(* IEC 61131-3 sources: daoli-st-library/DL_Motion (part 23) *)

(* ---- FB_DL_GantrySyncAxis.st ---- *)
(*==============================================================================
 * 组件名称 (Component)  : FB_DL_GantrySyncAxis
 * 所属子库 (Sublibrary) : DL_Motion
 * 当前版本 (Version)    : 1.0.0
 * 组件分类 (Category)   : 功能块（FUNCTION_BLOCK）· 多轴同步耦合族 · 龙门双驱偏斜保护
 * 兼容性   (Platform)   : CODESYS 3.5 / TwinCAT 3 / 汇川 InoProShop / Schneider
 *                         Machine Expert；仅依赖 Standard.library
 *                         （TON / R_TRIG / LIMIT / MIN / MAX / ABS），零厂商方言
 * 接口依赖 (Depends)    : I_DL_MotionAxis / E_DL_AxisState（既有契约，Round 05，零修改）
 * 功能描述 (Function)   : 双驱龙门同步与偏斜保护。主动侧（主轴）与从动侧（从轴）
 *                         1:1 速度耦合，实时监视两侧实际位置偏差；两级阈值（预警
 *                         / 故障）分别触发降速纠偏与双轴停止；可选比例纠偏（偏差
 *                         为正即主动侧在前 → 从动侧加速追赶）；任一轴故障同拍双轴
 *                         停止（不对称风险优先，不做「健康侧继续」策略）。
 * 设计要点 (Key notes)  :
 *   ① 两级监视是本块骨架：预警阈只告警与纠偏，故障阈才双停；预警阈必须小于
 *      故障阈，组态写反时自动对调并提示（沿用库内对调自修复先例）。
 *   ② 偏差确认走延时（抗单拍毛刺）；延时参数变化时显式断输入一拍，使已计时
 *      归零（防「改时间常数后计时不清零」的幽灵故障）。
 *   ③ 纠偏为比例律 + 修正量限幅，不用积分（避免在轴外层再套积分器造成饱和）；
 *      长时间饱和判为机械卡滞或增益不足，升为故障级锁存。
 *   ④ 偏差回差 80% 才退出纠偏态，防止阈值边缘反复抖动。
 * 开源溯源 (Origin)     : 原创实现，clean-room。语义来源为公开技术文章「双编码器
 *                         龙门组态」（两级位置差监视、偏差锁存门限）、公开厂商
 *                         帮助的软龙门章节（两级监视：一级可复位、二级不可复位）、
 *                         公开论文「宽跨距龙门吊防偏斜控制器」（偏差 → 速度修正
 *                         量、增益限幅）与公开的数控龙门位置公差参考值（来源编号
 *                         RAW_NOTES S-3）。
 *                         「借鉴对象的许可说明」：上述对象均为公开发布但受版权
 *                         保护的帮助文档 / 技术文章 / 公开论文，属「可免费查阅、
 *                         仅借鉴语义与参数域」类别；本实现未复制任何源码或组态
 *                         文件，状态机、引脚命名、故障码与对调自修复策略均为本
 *                         库自有设计。
 * 验收向量 (Acceptance) :
 *   V1 正常耦合：使能后进入 eRun，偏差在预警阈内 → bInSync 为 TRUE；
 *   V2 注入 1 mm 偏差：进入 eCorrecting，修正量不超上限，偏差收敛后回 eRun；
 *   V3 偏差 3 mm（超故障阈 2 mm）持续 60 ms：确认后双轴同时停止 + 锁存 0273；
 *   V4 单轴故障：同拍双轴停止 + 锁存 0274（不等待偏差阈值）；
 *   V5 阈值写反（预警 5 / 故障 1）：自动对调 + 信息级 0151，仍能正常监视；
 *   V6 纠偏饱和持续 3 s：锁存 0271；
 *   V7 偏差未回到预警阈内给 bReset：拒绝复位 + 信息级 0150；
 *   V8 位置含非有限值：锁存 0272 并立即双停；
 *   V9 运行中途插入跟踪脉冲 bTrack：清偏差计时、退回 eIdle（公约 0.1）。
 * 已知限制 (Limits)     :
 *   ① 本块为逻辑层同步监视与纠偏编排，不构成 ISO 13849 / IEC 62061 认证安全
 *      功能；机械偏斜的最终保护由硬件限位与安全回路承担。
 *   ② 两侧轴若注入同一实例，块内无法识别，轴自身仲裁；调用方须保证主动侧与
 *      从动侧为不同实例。
 *   ③ 偏差延时确认粒度等于任务扫描周期，极短延时（小于两个扫描周期）实际等效
 *      单拍确认，毛刺风险由调用方通过 tDevDelay 规避。
 * 规格偏离 (Deviation)  :
 *   ① 依公约 0.1 增补 bTrack 输入引脚（首扫 / 跟踪范式强制项）。
 *   ② 进入 eStopping 后沿用本块既有的停止单发标志，避免每拍重复下发停止指令；
 *      规格「同拍对两轴各发一次」在进入该态的同一拍内完成，语义不变。
 *   ③ 使能撤除时在清零输出的同时补发一次双轴停止（安全保守处置）。
 *   ④ 故障级码 0270（阈值非法）在使能期间逐拍复核，一旦组态被改坏立即锁存，
 *      不停留在仅启动时校验。
 * 红线自检 (Redline)    :
 *   R1 零全局符号区访问 ✓（无全局变量表访问、无外部变量声明）
 *   R2 零物理地址直写 ✓（无输入输出通道地址记号）
 *   R3 纯 IEC 61131-3 ✓（仅 TON / R_TRIG / LIMIT / MIN / MAX / ABS）
 *   R4 防除零 / 防越界 / 浮点容差 ✓（阈值对调与回差全用容差比较、无数组索引、
 *      时间参数变化断输入一拍）
 *   R5 声明行 100% 中英双语同行注释 ✓
 *   R6 ENUM + CASE 且 CASE 含 ELSE 兜底 ✓
 *   R7 定时器与边沿实例无条件周期刷新 ✓（本块无单拍脉冲输出）
 *   POU 终结符成对 ✓（FUNCTION_BLOCK ↔ END_FUNCTION_BLOCK，末行即终结符；
 *   TYPE ↔ END_TYPE 成对）
 * 故障码表 (Error codes):
 *   16#0004_0150【信息级】偏差未回预警阈内，复位被拒；
 *   16#0004_0151【信息级】预警 / 故障阈值对调自修复；
 *   16#0004_0152【信息级】纠偏速度上限非法回默认；
 *   16#0004_0270【故障级】偏差阈值非法（≤0 / 非有限值），锁存；
 *   16#0004_0271【故障级】纠偏长时间饱和（疑似机械卡滞），锁存；
 *   16#0004_0272【故障级】轴位置信号非有限值，锁存；
 *   16#0004_0273【故障级】偏差超故障阈触发双轴停止，锁存；
 *   16#0004_0274【故障级】单轴故障触发双轴停止（透传），锁存；
 *   16#0004_0297【故障级】非法状态兜底（本块专用，不与其他块共用）。
 *   信息级码只进 uErrorId；bFault 为派生式仅反映 eFault 态。
 * 修订历史 (Revision)   :
 *   2026-11-15  v1.0.0  首版入库（Round 08 · DL_Motion 同步耦合族）
 *============================================================================*)

(*-----------------------------------------------------------------------------
 * 调用示例 (Instance guide)：
 *   fbGantry.iMasterAxis := fbLeftAxis;           // 主动侧（驱动侧）实例
 *   fbGantry.iSlaveAxis  := fbRightAxis;          // 从动侧（跟随侧）实例
 *   fbGantry(bEnable := bGantryOn,
 *            fDevTolWarn := 0.5, fDevTolFault := 2.0,
 *            tDevDelay := T#50MS, bCorrectEnable := TRUE,
 *            fCorrGain := 2.0, fCorrSpeedMax := 20.0,
 *            fCoupleSpeed := 10.0, fAcc := 500.0);
 *   IF fbGantry.bStopBothCmd THEN bSafetyRelayDrop := TRUE; END_IF
 *   注：两侧轴的上使能、回原与限位保护仍由各自轴块与安全链负责，本块只做
 *       速度耦合与偏差监视。
 *----------------------------------------------------------------------------*)

(*-----------------------------------------------------------------------------
 * 常见误用与现场提示 (Field notes)：
 *   1 预警阈与故障阈不要设成同值：同值时监视失去两级意义，块内会按对调处理
 *      并提示，但工艺上应重新组态（预警阈建议取故障阈的 1/4 ~ 1/2）。
 *   2 纠偏增益过大会在阈值边缘产生速度抖动；从 1.0 ~ 3.0 起步，观察
 *      fCorrSpeedCmd 是否长期贴上限（贴上限即增益不足或机械卡滞）。
 *   3 单轴报跟随误差时本块同拍双停，另一轴不会「继续跑」——这是刻意的保守
 *      策略，复位后必须人工确认横梁已回正再重新使能。
 *   4 bFault 一旦置位只能靠 bReset 上升沿解除，且要求偏差已回到预警阈内；
 *      机械偏斜未消除时复位会被拒（信息级 0150），必须先手动点动纠偏。
 *   5 本块不产生位置指令，只产生速度指令；位置同步精度取决于两侧驱动自身
 *      的位置环，本块不替代驱动的位置控制。
 *   6 阈值组态被改坏（≤0 / 非有限值 / 超域）时本块直接锁存 0270，且「组态未改好
 *      之前复位会立刻再次锁存」是刻意行为：不允许带着非法偏差阈值运行龙门。
 *----------------------------------------------------------------------------*)

(*-----------------------------------------------------------------------------
 * 枚举: E_DL_GantryState（归属 DL_Motion，与本功能块同文件发布）
 * 含义: 龙门双驱同步状态机，编号间隔 10 预留扩展位。
 *----------------------------------------------------------------------------*)
{attribute 'strict'}
{attribute 'qualified_only'}
TYPE E_DL_GantryState :
(
    eIdle       := 0,    // 空闲：未耦合，输出全清 / Idle: not coupled, outputs cleared
    eCoupling   := 10,   // 耦合建立：双轴以慢速趋同 / Coupling: both axes converge at low speed
    eRun        := 20,   // 运行：1:1 速度跟随 + 偏差监视 / Run: 1:1 velocity follow with deviation monitoring
    eCorrecting := 30,   // 纠偏中：偏差超预警阈且纠偏使能 / Correcting: deviation over warn band with correction enabled
    eStopping   := 40,   // 双轴停止中：偏差超故障阈或任一轴故障 / Stopping: deviation over fault band or axis fault
    eFault      := 99    // 故障锁存：仅 bReset 上升沿且偏差回位可退出 / Fault: latched, bReset only after deviation recovered
) UINT;
END_TYPE

FUNCTION_BLOCK FB_DL_GantrySyncAxis
VAR_INPUT
    bEnable         : BOOL := FALSE;        // 总使能（Enable），FALSE=停止并清指令，电平语义
    bReset          : BOOL := FALSE;        // 复位故障（Reset），上升沿受理，须偏差已回预警阈内才真正复位
    bTrack          : BOOL := FALSE;        // 偏差计时重同步（Tracking pulse），上升沿即清计时与锁存并退回 eIdle
    fDevTolWarn     : REAL := 0.5;          // 偏差预警阈（Deviation warn tolerance）[mm]，域 0.001..50，须小于故障阈
    fDevTolFault    : REAL := 2.0;          // 偏差故障阈（Deviation fault tolerance）[mm]，域 0.01..100
    tDevDelay       : TIME := T#50MS;       // 偏差确认延时（Deviation confirm delay）[ms]，超阈须持续此时间才动作
    bCorrectEnable  : BOOL := TRUE;         // 纠偏使能（Correction enable），FALSE=只监视不纠偏
    fCorrGain       : REAL := 2.0;          // 纠偏比例增益（Correction gain）[1/s]，域 0..50，0=纠偏关闭
    fCorrSpeedMax   : REAL := 20.0;         // 纠偏速度修正上限（Correction speed limit）[mm/s]，域 0.1..500
    fCoupleSpeed    : REAL := 10.0;         // 耦合建立慢速（Coupling speed）[mm/s]，域 0.1..1000，双轴以此速度趋同
    fAcc            : REAL := 500.0;        // 加/减速度（Acceleration）[mm/s²]，域 0.1..100000，非有限值回默认
END_VAR
VAR_OUTPUT
    bInSync         : BOOL := FALSE;        // 同步中（In sync），eRun / eCorrecting 且偏差未超预警阈为 TRUE
    fDeviation      : REAL := 0.0;          // 实时偏差（Deviation）[mm]，= 主动侧位置 − 从动侧位置，带符号
    bDevWarn        : BOOL := FALSE;        // 偏差预警（Deviation warning），延时确认后置位，回差内自动清，瞬态型
    bFault          : BOOL := FALSE;        // 故障锁存（Fault），派生式仅故障级码参与，信息级码不置位
    uErrorId        : UDINT := 0;           // 故障码（Error code），段位 16#0004_xxxx，0=无故障
    bStopBothCmd    : BOOL := FALSE;        // 双轴停止请求（Stop both request），供上层安全链与 HMI 监视
    fCorrSpeedCmd   : REAL := 0.0;          // 纠偏速度修正量（Correction speed）[mm/s]，带符号，叠加到从动侧指令
END_VAR
VAR_IN_OUT
    iMasterAxis     : I_DL_MotionAxis;      // 主动侧轴接口引用（Drive side axis），由调用方注入
    iSlaveAxis      : I_DL_MotionAxis;      // 从动侧轴接口引用（Following side axis），由调用方注入
END_VAR
VAR
    eState          : E_DL_GantryState := E_DL_GantryState.eIdle; // 内部状态机步序（Internal state）
    bInit           : BOOL := FALSE;        // 首扫完成标志（First-scan done flag），初值 FALSE，随 bTrack 复位
    bFaultLatch     : BOOL := FALSE;        // 故障锁存标志（Fault latch），仅 bReset 沿或新啮合沿解除
    bRefOk          : BOOL := FALSE;        // 双引用有效标志（Both references valid），逐拍重算
    bStopIssued     : BOOL := FALSE;        // 双轴停止已下发标志（Stop issued flag），单发化防重复发令
    bWarnLatched    : BOOL := FALSE;        // 预警锁存标志（Warning latched），带回差自动清除
    bMonActive      : BOOL := FALSE;        // 偏差监视使能（Monitoring active），运行三态为 TRUE
    bParamBad       : BOOL := FALSE;        // 阈值参数非法标志（Tolerance parameter invalid），逐拍重算
    bDelayChanged   : BOOL := FALSE;        // 延时参数变更标志（Delay changed flag），断输入一拍用
    fWarnEff        : REAL := 0.5;          // 生效预警阈（Effective warn tolerance）[mm]，对调后值
    fFaultEff       : REAL := 2.0;          // 生效故障阈（Effective fault tolerance）[mm]，对调后值
    fCorrMaxEff     : REAL := 20.0;         // 生效纠偏上限（Effective correction limit）[mm/s]，非法回默认
    fAccEff         : REAL := 500.0;        // 生效加减速度（Effective acceleration）[mm/s²]，非法回默认
    fCoupleEff      : REAL := 10.0;         // 生效耦合慢速（Effective coupling speed）[mm/s]，非法回默认
    fDevAbs         : REAL := 0.0;          // 偏差绝对值（Absolute deviation）[mm]，阈值比较用
    fCorrAbs        : REAL := 0.0;          // 纠偏量绝对值（Absolute correction）[mm/s]，饱和判定用
    fCorrCmd        : REAL := 0.0;          // 纠偏修正量（Correction command）[mm/s]，带符号
    fMasterPos      : REAL := 0.0;          // 主动侧位置（Drive side position）[mm]
    fSlavePos       : REAL := 0.0;          // 从动侧位置（Following side position）[mm]
    fMasterVel      : REAL := 0.0;          // 主动侧速度（Drive side velocity）[mm/s]，带符号
    fSlaveVel       : REAL := 0.0;          // 从动侧速度（Following side velocity）[mm/s]，带符号
    fCmdVel         : REAL := 0.0;          // 下发给从动侧的速度指令（Commanded velocity）[mm/s]，带符号
    tDelayEff       : TIME := T#50MS;       // 生效确认延时（Effective confirm delay）[ms]，负值归零
    tDelayPrev      : TIME := T#0MS;        // 上拍确认延时（Previous confirm delay）[ms]，变更检测基准
    nStopCode       : UDINT := 0;           // 停止原因码（Stop reason code），进 eFault 时落地
    fbTrigReset     : R_TRIG;               // 复位指令上升沿（Reset command rising edge）
    fbTonDevWarn    : TON;                  // 偏差预警延时确认（Warn confirm delay timer）
    fbTonDevFault   : TON;                  // 偏差故障延时确认（Fault confirm delay timer）
    fbTonCorrSat    : TON;                  // 纠偏饱和累计计时（Correction saturation timer）
END_VAR
VAR CONSTANT
    DL_GANTRY_INF_MAX   : REAL := 1.0E30;   // 有限值判定幅值上限（Finite magnitude bound）[无量纲，按比较量量纲同值使用]
    DL_GANTRY_EPS       : REAL := 1.0E-6;   // 浮点判零容差（Float zero tolerance）[无量纲，按比较量量纲同值使用]
    DL_GANTRY_TOL_MIN   : REAL := 1.0E-3;   // 阈值下限（Tolerance floor）[mm]，低于此值判非法
    DL_GANTRY_TOL_MAX   : REAL := 100.0;    // 阈值上限（Tolerance ceiling）[mm]，高于此值判非法
    DL_GANTRY_CORR_DEF  : REAL := 20.0;     // 纠偏上限默认值（Default correction limit）[mm/s]
    DL_GANTRY_CORR_MAX  : REAL := 500.0;    // 纠偏上限允许最大值（Correction limit ceiling）[mm/s]
    DL_GANTRY_ACC_DEF   : REAL := 500.0;    // 加速度默认回退值（Default acceleration）[mm/s²]
    DL_GANTRY_CPL_DEF   : REAL := 10.0;     // 耦合慢速默认回退值（Default coupling speed）[mm/s]
    DL_GANTRY_HYST      : REAL := 0.8;      // 回差系数（Hysteresis factor）[-]，低于预警阈 80% 才清预警
    DL_GANTRY_SAT_RATIO : REAL := 0.98;     // 饱和判定比例（Saturation ratio）[-]，达上限 98% 视为饱和
    DL_GANTRY_SAT_TIME  : TIME := T#3S;     // 饱和持续上限（Saturation time limit）[ms]，超过判卡滞
    DL_GANTRY_SPEED_BAND: REAL := 1.0E-5;   // 速度趋同判定带（Speed convergence band）[mm/s]，= 判零容差 × 10
    DL_GANTRY_ZERO_TIME : TIME := T#0S;     // 零延时字面量（Zero delay literal）[ms]，用于延时下限比较
END_VAR

// 段 1｜边沿实例无条件周期刷新（红线 R7：严禁置于 IF / CASE 分支内）
fbTrigReset(CLK := bReset);

// 段 2｜出口默认赋值（公约 0.9：早退路径输出必须确定）
bInSync       := FALSE;
bDevWarn      := FALSE;
bFault        := (eState = E_DL_GantryState.eFault);
fCorrSpeedCmd := 0.0;
fDeviation    := 0.0;

// 段 3｜双引用有效性判定 + 反馈量采集（无效时全部回零，定时器照样刷新）
bRefOk := (iMasterAxis <> 0) AND (iSlaveAxis <> 0);
IF bRefOk THEN
    fMasterPos := iMasterAxis.fPosition;
    fSlavePos  := iSlaveAxis.fPosition;
    fMasterVel := iMasterAxis.fVelocity;
    fSlaveVel  := iSlaveAxis.fVelocity;
ELSE
    fMasterPos := 0.0;
    fSlavePos  := 0.0;
    fMasterVel := 0.0;
    fSlaveVel  := 0.0;
END_IF
fDeviation := fMasterPos - fSlavePos;
fDevAbs    := ABS(fDeviation);

// 段 4｜阈值参数防御：非有限值 / 超域判非法，预警阈不小于故障阈时自动对调
fWarnEff  := fDevTolWarn;
fFaultEff := fDevTolFault;
bParamBad := FALSE;
IF (fWarnEff <> fWarnEff) OR (ABS(fWarnEff) > DL_GANTRY_INF_MAX)
   OR (fWarnEff < DL_GANTRY_TOL_MIN) OR (fWarnEff > DL_GANTRY_TOL_MAX) THEN
    bParamBad := TRUE;
END_IF
IF (fFaultEff <> fFaultEff) OR (ABS(fFaultEff) > DL_GANTRY_INF_MAX)
   OR (fFaultEff < DL_GANTRY_TOL_MIN) OR (fFaultEff > DL_GANTRY_TOL_MAX) THEN
    bParamBad := TRUE;
END_IF
IF (NOT bParamBad) AND (fWarnEff > (fFaultEff - DL_GANTRY_EPS)) THEN
    fWarnEff  := fDevTolFault;                           // 自动对调：写反时按对调后值监视，不静默
    fFaultEff := fDevTolWarn;
    uErrorId  := 16#0004_0151;                           // 【信息级】预警 / 故障阈值对调自修复
END_IF

IF (fCorrSpeedMax <> fCorrSpeedMax) OR (ABS(fCorrSpeedMax) > DL_GANTRY_INF_MAX)
   OR (fCorrSpeedMax < DL_GANTRY_TOL_MIN) THEN
    fCorrMaxEff := DL_GANTRY_CORR_DEF;                   // 纠偏上限非法 → 默认 20 mm/s
    uErrorId    := 16#0004_0152;                         // 【信息级】纠偏速度上限非法回默认
ELSE
    fCorrMaxEff := MIN(fCorrSpeedMax, DL_GANTRY_CORR_MAX);
END_IF

IF (fAcc <> fAcc) OR (ABS(fAcc) > DL_GANTRY_INF_MAX) OR (fAcc < DL_GANTRY_TOL_MIN) THEN
    fAccEff := DL_GANTRY_ACC_DEF;
ELSE
    fAccEff := fAcc;
END_IF

IF (fCoupleSpeed <> fCoupleSpeed) OR (ABS(fCoupleSpeed) > DL_GANTRY_INF_MAX) OR (fCoupleSpeed < DL_GANTRY_TOL_MIN) THEN
    fCoupleEff := DL_GANTRY_CPL_DEF;
ELSE
    fCoupleEff := fCoupleSpeed;
END_IF

// 段 5｜确认延时防御与变更检测（公约 0.6：语义参数变化必须断输入一拍）
IF tDevDelay < DL_GANTRY_ZERO_TIME THEN
    tDelayEff := DL_GANTRY_ZERO_TIME;                    // 负延时归零，按单拍确认（毛刺风险由调用方规避）
ELSE
    tDelayEff := tDevDelay;
END_IF
bDelayChanged := (tDelayEff <> tDelayPrev);              // 延时变更：本拍强制断输入，使已计时归零
tDelayPrev    := tDelayEff;

// 段 6｜偏差监视使能（运行三态参与监视）
bMonActive := (eState = E_DL_GantryState.eCoupling) OR (eState = E_DL_GantryState.eRun)
              OR (eState = E_DL_GantryState.eCorrecting);

// 段 7｜定时器无条件周期刷新（红线 R7：严禁置于 IF / CASE 分支内）
fbTonDevWarn(IN := bRefOk AND bMonActive AND (fDevAbs >= fWarnEff) AND (NOT bDelayChanged),
             PT := tDelayEff);
fbTonDevFault(IN := bRefOk AND bMonActive AND (fDevAbs >= fFaultEff) AND (NOT bDelayChanged),
              PT := tDelayEff);
fbTonCorrSat(IN := (eState = E_DL_GantryState.eCorrecting) AND (fCorrAbs >= fCorrMaxEff * DL_GANTRY_SAT_RATIO),
             PT := DL_GANTRY_SAT_TIME);

// 段 8｜引用无效直接退出（定时器已在上方无条件刷新，本拍不产生任何轴动作）
IF NOT bRefOk THEN
    RETURN;
END_IF

// 段 9｜预警锁存与回差清除（瞬态型，每拍重算）
IF fDevAbs >= fWarnEff THEN
    bWarnLatched := fbTonDevWarn.Q;                      // 超阈值区间：以延时确认结果为准
ELSIF fDevAbs <= (fWarnEff * DL_GANTRY_HYST) THEN
    bWarnLatched := FALSE;                               // 回差内自动清除
END_IF

// 段 10｜首扫与跟踪范式（公约 0.1：bTrack OR (NOT bInit) 为唯一判据，禁止反序）
IF bTrack OR (NOT bInit) THEN
    bWarnLatched := FALSE;
    bStopIssued  := FALSE;
    bStopBothCmd := FALSE;
    fCorrCmd     := 0.0;
    fCorrAbs     := 0.0;
    nStopCode    := 0;
    eState       := E_DL_GantryState.eIdle;
    bInit        := TRUE;                                // 首扫完成后置位（判据恒为 bTrack OR NOT bInit）
END_IF

// 段 11｜总使能撤除：清指令 + 补发一次双轴停止（安全保守处置）
IF NOT bEnable THEN
    IF (NOT bStopIssued) AND ((eState = E_DL_GantryState.eCoupling) OR (eState = E_DL_GantryState.eRun)
       OR (eState = E_DL_GantryState.eCorrecting)) THEN
        iMasterAxis.Stop();                              // 主动侧停止（本拍唯一一次主动侧调用）
        iSlaveAxis.Stop();                               // 从动侧停止（本拍唯一一次从动侧调用）
        bStopIssued := TRUE;
    END_IF
    eState    := E_DL_GantryState.eIdle;
    fCorrCmd  := 0.0;
    fCorrAbs  := 0.0;
END_IF

// 段 12｜事件码管理（公约 0.7 / R15）：锁存码仅在解除路径清，瞬时码逐拍重算
IF NOT bFaultLatch THEN
    uErrorId := 0;
END_IF

// 段 13｜位置 / 力矩类信号非有限值拦截（判定不可信，立即转双停）
IF (fMasterPos <> fMasterPos) OR (fSlavePos <> fSlavePos)
   OR (ABS(fMasterPos) > DL_GANTRY_INF_MAX) OR (ABS(fSlavePos) > DL_GANTRY_INF_MAX) THEN
    IF (eState <> E_DL_GantryState.eIdle) AND (eState <> E_DL_GantryState.eFault) THEN
        nStopCode := 16#0004_0272;                       // 【故障级】轴位置信号非有限值
        eState    := E_DL_GantryState.eStopping;
    END_IF
END_IF

// 段 14｜阈值非法拦截（使能期间逐拍复核组态）
IF bParamBad THEN
    IF eState <> E_DL_GantryState.eFault THEN
        bFaultLatch := TRUE;
        uErrorId    := 16#0004_0270;                     // 【故障级】偏差阈值非法
        eState      := E_DL_GantryState.eFault;
    END_IF
END_IF

// 段 15｜主状态机（ENUM + CASE + ELSE 兜底）
CASE eState OF

    E_DL_GantryState.eIdle:                              // 空闲：等待使能
        bInSync  := FALSE;
        bStopIssued := FALSE;
        bStopBothCmd := FALSE;
        fCorrCmd := 0.0;
        IF bEnable AND (NOT bParamBad) THEN
            bFaultLatch := FALSE;                        // 使能上升：锁存码解除路径（R15）
            fCorrCmd    := 0.0;
            eState      := E_DL_GantryState.eCoupling;
        END_IF

    E_DL_GantryState.eCoupling:                          // 耦合建立：双轴以慢速趋同
        bStopBothCmd := FALSE;
        IF iMasterAxis.bError OR iSlaveAxis.bError THEN
            nStopCode := 16#0004_0274;                   // 【故障级】单轴故障（不对称风险优先）
            eState    := E_DL_GantryState.eStopping;
        ELSIF fbTonDevFault.Q THEN
            nStopCode := 16#0004_0273;                   // 【故障级】偏差超故障阈
            eState    := E_DL_GantryState.eStopping;
        ELSE
            // 跟随主动侧速度，但幅值不超过耦合慢速
            fCmdVel := LIMIT(-fCoupleEff, fMasterVel, fCoupleEff);
            IF NOT iSlaveAxis.MoveVelocity(fVel := fCmdVel, fAcc := fAccEff) THEN
                bFaultLatch := TRUE;
                uErrorId    := 16#0004_0274;             // 【故障级】从动侧速度指令被拒（按单轴故障处置）
                eState      := E_DL_GantryState.eFault;
            ELSIF (ABS(fMasterVel - fSlaveVel) <= DL_GANTRY_SPEED_BAND) AND (fDevAbs <= fWarnEff) THEN
                eState := E_DL_GantryState.eRun;         // 速度趋同且偏差在预警阈内 → 运行
            END_IF
        END_IF

    E_DL_GantryState.eRun:                               // 运行：1:1 跟随，纠偏量为零
        IF iMasterAxis.bError OR iSlaveAxis.bError THEN
            nStopCode := 16#0004_0274;
            eState    := E_DL_GantryState.eStopping;
        ELSIF fbTonDevFault.Q THEN
            nStopCode := 16#0004_0273;
            eState    := E_DL_GantryState.eStopping;
        ELSE
            fCorrCmd := 0.0;                             // 运行态不纠偏
            IF bCorrectEnable AND (ABS(fCorrGain) > DL_GANTRY_EPS) AND bWarnLatched THEN
                eState := E_DL_GantryState.eCorrecting;  // 偏差确认超预警阈且纠偏使能 → 纠偏
            END_IF
            fCmdVel := fMasterVel;
            IF NOT iSlaveAxis.MoveVelocity(fVel := fCmdVel, fAcc := fAccEff) THEN
                bFaultLatch := TRUE;
                uErrorId    := 16#0004_0274;             // 【故障级】从动侧速度指令被拒
                eState      := E_DL_GantryState.eFault;
            END_IF
        END_IF

    E_DL_GantryState.eCorrecting:                        // 纠偏中：比例律修正量限幅
        IF iMasterAxis.bError OR iSlaveAxis.bError THEN
            nStopCode := 16#0004_0274;
            eState    := E_DL_GantryState.eStopping;
        ELSIF fbTonDevFault.Q THEN
            nStopCode := 16#0004_0273;
            eState    := E_DL_GantryState.eStopping;
        ELSIF fbTonCorrSat.Q THEN
            bFaultLatch := TRUE;
            uErrorId    := 16#0004_0271;                 // 【故障级】纠偏长时间饱和（疑似卡滞 / 增益不足）
            eState      := E_DL_GantryState.eFault;
        ELSE
            // 偏差为正（主动侧在前）→ 从动侧加速追赶；为负则减速
            fCorrCmd := LIMIT(-fCorrMaxEff, fCorrGain * fDeviation, fCorrMaxEff);
            fCorrAbs := ABS(fCorrCmd);
            // 偏差回到预警阈 80% 以内（回差）→ 退出纠偏
            IF fDevAbs <= (fWarnEff * DL_GANTRY_HYST) THEN
                fCorrCmd := 0.0;
                fCorrAbs := 0.0;
                eState   := E_DL_GantryState.eRun;
            END_IF
            fCmdVel := fMasterVel + fCorrCmd;
            IF NOT iSlaveAxis.MoveVelocity(fVel := fCmdVel, fAcc := fAccEff) THEN
                bFaultLatch := TRUE;
                uErrorId    := 16#0004_0274;             // 【故障级】从动侧速度指令被拒
                eState      := E_DL_GantryState.eFault;
            END_IF
        END_IF

    E_DL_GantryState.eStopping:                          // 双轴停止：同拍各发一次，停稳后锁存
        bStopBothCmd := TRUE;
        fCorrCmd     := 0.0;
        fCorrAbs     := 0.0;
        IF NOT bStopIssued THEN
            iMasterAxis.Stop();                          // 主动侧停止（本拍唯一一次主动侧调用）
            iSlaveAxis.Stop();                           // 从动侧停止（本拍唯一一次从动侧调用）
            bStopIssued := TRUE;
        END_IF
        IF (ABS(fMasterVel) <= DL_GANTRY_EPS) AND (ABS(fSlaveVel) <= DL_GANTRY_EPS) THEN
            bFaultLatch := TRUE;
            IF nStopCode = 0 THEN
                uErrorId := 16#0004_0273;                // 【故障级】兜底：停止原因缺失时按偏差超限记账
            ELSE
                uErrorId := nStopCode;                   // 落地本次停止的真实原因码
            END_IF
            bStopIssued := FALSE;
            eState      := E_DL_GantryState.eFault;
        END_IF

    E_DL_GantryState.eFault:                             // 故障锁存：仅复位沿且偏差回位可退出
        bInSync      := FALSE;
        bStopBothCmd := TRUE;                            // 故障态保持停止请求，供安全链与 HMI 监视
        fCorrCmd     := 0.0;
        fCorrAbs     := 0.0;
        bStopIssued  := FALSE;
        IF fbTrigReset.Q THEN
            IF fDevAbs <= fWarnEff THEN
                bFaultLatch := FALSE;                    // 唯一解除路径：偏差已回预警阈内
                uErrorId    := 0;
                nStopCode   := 0;
                eState      := E_DL_GantryState.eIdle;
            ELSE
                uErrorId := 16#0004_0150;                // 【信息级】偏差未回预警阈内，复位被拒
            END_IF
        END_IF

    ELSE                                                 // 非法状态兜底（本块专用码）
        bFaultLatch  := TRUE;
        uErrorId     := 16#0004_0297;                    // 【故障级】非法状态兜底
        bInSync      := FALSE;
        bStopBothCmd := TRUE;
        fCorrCmd     := 0.0;
        fCorrAbs     := 0.0;
        eState       := E_DL_GantryState.eFault;

END_CASE

// 段 16｜出口映射（派生式，信息级码不参与 bFault）
bFault        := (eState = E_DL_GantryState.eFault);
bInSync       := ((eState = E_DL_GantryState.eRun) OR (eState = E_DL_GantryState.eCorrecting))
                 AND (NOT bWarnLatched);
bDevWarn      := bWarnLatched AND ((eState = E_DL_GantryState.eCoupling)
                 OR (eState = E_DL_GantryState.eRun) OR (eState = E_DL_GantryState.eCorrecting));
bStopBothCmd  := (eState = E_DL_GantryState.eStopping) OR (eState = E_DL_GantryState.eFault);
fDeviation    := fMasterPos - fSlavePos;
fCorrSpeedCmd := fCorrCmd;

END_FUNCTION_BLOCK

(* ---- FB_DL_LineInterp2Axis.st ---- *)
(*==============================================================================
 * 组件名称 (Component)  : FB_DL_LineInterp2Axis
 * 所属子库 (Sublibrary) : DL_Motion
 * 当前版本 (Version)    : 1.0.1
 * 组件分类 (Category)   : 功能块（FUNCTION_BLOCK）· 运动控制 · 两轴直线插补
 * 兼容性   (Platform)   : CODESYS 3.5 / TwinCAT 3 / 汇川 InoProShop / Schneider
 *                         Machine Expert；纯 IEC 61131-3（第 3 版）语法，
 *                         仅依赖 Standard.library（R_TRIG / SQRT / MIN / MAX / LIMIT）
 * 功能描述 (Function)   : 由起点、终点、合成速度与加速度生成两轴位置给定：单位向量分解、
 *                         单轴速度上限折算、梯形与三角速度曲线自适应、端点平滑减速、
 *                         暂停保持与故障保护。输出 X 与 Y 的位置给定、合成速度、完成度
 *                         与本次实际峰值速度。
 * 分层声明 (Layering)   : ① 本件只输出「位置给定」，不输出使能、回零与报警复位，也不直接
 *                         驱动物理轴——两轴的实际闭环由各自的单轴功能块承担，本件给出
 *                         给定值后由上层把给定接到单轴的相对或绝对运动接口；
 *                         ② 不读系统时钟、不读任务周期：插补时间增量由引脚注入，
 *                         保证结果可复现、跨平台一致；
 *                         ③ 不做圆弧与样条插补（属后续件），不做过象限与软限位判断
 *                         （软限位归运动层的软限位保护件）。
 * 周期纪律 (Cycle)      : 本件必须放在固定周期任务中调用，周期值通过标称周期引脚注入。
 *                         变周期任务（如带事件触发的任务）会直接造成速度与位置偏差，
 *                         因为时间增量按注入值推进、不按墙钟补偿。
 * 速度剖面 (Profile)    : 单侧加速度距离为合成速度平方除以两倍加速度；若两侧之和超过
 *                         路径总长则判为三角曲线，峰值速度降为「加速度乘路径长」的平方根，
 *                         加速距离取路径长的一半。临界相等（两侧之和恰等于路径长）按梯形
 *                         处理：此时峰值速度与期望合成速度相等，两种判法结果一致、不跳变。
 * 端点纪律 (Endpoint)   : 减速段出口强制把已走距离钳到路径总长，进度置 100，避免离散步长
 *                         越过终点导致给定超程；收尾速度保留峰值的若干比例，防止速度
 *                         指数衰减而出现「永远差最后一点」的爬行。
 * 开源溯源 (Origin)     : 来源标签 github-topics-motion。原创实现（参考 GitHub 运动控制与
 *                         结构化文本主题下开源运动库的共同形态：单位向量分解、合成速度
 *                         限幅、梯形与三角自适应三段结构；多份实现交叉印证其为社区共识
 *                         写法，非某一家独有）。速度剖面、临界判据、暂停策略、枚举、
 *                         状态机与全部码位 100% 本库独立设计，clean-room 实现，零代码行
 *                         复制。各上游仓库许可未逐条复核，按最严口径只借结构与参数域。
 * 依赖     (Depends)    : 无 DL_ 内部依赖；Standard.library: R_TRIG / SQRT / MIN / MAX / LIMIT
 * 故障码表 (Error codes):
 *   16#0004_0109【信息级】路径长度为零，当拍直接完成，给定等于起点
 *   16#0004_010A【信息级】标称周期越界已钳到 0.1 毫秒至 1 秒
 *   16#0004_010B【信息级】单轴速度上限参与折算，合成速度已被压低
 *   16#0004_010C【信息级】路径过短，速度曲线降为三角（无匀速段）
 *   16#0004_0204【故障级】速度、加速度、单轴限速或最大路径长参数非法（锁存）
 *   16#0004_0205【故障级】路径长度超过允许上限（锁存）
 *   16#0004_0206【故障级】输入含非有限值（NaN 或无穷），前置拦截（锁存）
 *   16#0004_0207【故障级】非法状态兜底（锁存，终端安全态）
 * 码位占用 (Slot)       : 信息级 0109 / 010A / 010B / 010C；故障级 0204 / 0205 / 0206 / 0207。
 *                         全部落在 R12 本件分配块内，无跨块借用、无段外哨兵值。
 * 拍序纪律 (Cycle order) :
 *   ① ePhase    ：段 7 状态机（唯一位移点），段 8 复位分支是唯一回退点
 *   ② fS 与 fV  ：只在加速、匀速、减速三段内推进；暂停段速度归零且不推进位移
 *   ③ _bDone    ：进入准备相与进入完成相两处写，互斥不覆盖
 *   ④ uErrorId  ：段 9 单一优先级链，全拍只写一次
 * 验收向量 (Acceptance) :
 *   V1 梯形：起点 0 0、终点 300 400 → 路径 500；速度 100、加速度 200、单轴限速 1000 →
 *      合成 100 未被压低、单侧加速距离 25，两侧 50 小于 500 判梯形，峰值 100；
 *      中点给定为 150 与 200、完成度 50、合成速度 100
 *   V2 单轴限速：与 V1 同参但 X 轴限速改为 50 → 折算 83.333，合成速度被压到 83.333，
 *      X 分量 83.333 乘 0.6 等于 50，恰好不超限
 *   V3 零长度：起终点相同 → 当拍完成、给定等于起点、进度 100、码 0109
 *   V4 临界：路径 50、单侧加速距离 25 → 和为 50 恰等于路径长，判梯形，峰值 100
 *   V5 三角：路径 40 → 两侧 50 大于 40 判三角，峰值 89.44、单侧加速距离 20
 *   V6 参数非法：加速度为 0 → 故障位置位、码 0204、忙碌为假
 * 偏离留档 (Deviation)  :
 *   ① 规格未规定暂停时的时间补偿策略，本件按「不做补偿」实现：恢复后从当前速度重新加速，
 *      但时间增量仍按标称周期推进，故暂停不会造成位置瞬跳。若需要恒速衔接，应在工艺层
 *      用缓停而非暂停。
 *   ② 规格的减速段出口只要求钳位，本件额外把进度强制置 100，避免浮点除法在末拍给出
 *      99.9999 而让画面闪烁。
 * 修订历史 (Revision)   :
 *   2026-11-15  v1.0.0  首版落盘（R12 · 泳道 C · 两轴直线插补件）
 *   2026-11-15  v1.0.1  终审修复两处：
 *                       ① 暂停恢复时速度阶跃——加速段出口只看「位移到加速距离」，恢复后
 *                       该条件当拍即成立，再加速被整段跳过，速度由零直接跳到峰值；
 *                       改为位移与速度双条件，并在恢复时按剩余距离分流到减速段。
 *                       ② 零长度路径的完成度与头注释矛盾（注释写 100、出口被覆写为 0），
 *                       完成相下补满值分支
 *============================================================================*)

(*------------------------------------------------------------------------------
 * 枚举: E_DL_LineInterpPhase（本块相位，归属本功能块并同文件发布）
 *       Phase enumeration owned by this block, one member per motion segment
 *-----------------------------------------------------------------------------*)
TYPE E_DL_LineInterpPhase :
(
    eIdle  := 0,   // 待机：等待启动沿，给定保持在起点 / Idle, waiting for the start edge
    ePrep  := 10,  // 准备：参数闸门、向量分解、速度剖面计算 / Preparation, the whole profile is computed here
    eAccel := 20,  // 加速：速度按加速度上升，位移按速度积分 / Acceleration segment
    eCruise:= 30,  // 匀速：速度保持峰值，位移按速度积分 / Constant speed segment
    eDecel := 40,  // 减速：速度按加速度下降，出口钳位到终点 / Deceleration segment
    eDone  := 50,  // 完成：完成标志保持，给定等于终点，等下一次启动 / Done, held until the next start
    eHeld  := 60,  // 暂停：速度归零、位移保持，恢复后重新加速 / Held, speed forced to zero
    eFault := 99   // 故障：参数或输入非法、路径超限、非法状态 / Fault, needs a reset to leave
);
END_TYPE

FUNCTION_BLOCK FB_DL_LineInterp2Axis
VAR_INPUT
    bEnable       : BOOL;                          // 使能，FALSE 时停止推进并回待机 [-] / Enable, stopping the move and returning to idle
    bReset        : BOOL;                          // 复位故障，上升沿有效 [-] / Rising edge clears the fault
    bStart        : BOOL;                          // 启动，上升沿有效（待机与完成态可受理）[-] / Rising edge starts the move in idle or done
    bHold         : BOOL;                          // 暂停，TRUE 时速度归零且位移保持 [-] / Pauses the interpolation while TRUE
    fStartX       : REAL;                          // 起点 X 坐标 [毫米] / Start X in millimetres
    fStartY       : REAL;                          // 起点 Y 坐标 [毫米] / Start Y in millimetres
    fEndX         : REAL;                          // 终点 X 坐标 [毫米] / End X in millimetres
    fEndY         : REAL;                          // 终点 Y 坐标 [毫米] / End Y in millimetres
    fPathSpeed    : REAL := 100.0;                 // 期望合成速度 [毫米每秒]，域大于 0 / Desired path speed, must exceed zero
    fAccel        : REAL := 500.0;                 // 加减速度 [毫米每二次方秒]，域大于 0 / Acceleration, must exceed zero
    fMaxSpeedX    : REAL := 1000.0;                // X 轴速度上限 [毫米每秒]，域大于 0 / X axis speed limit
    fMaxSpeedY    : REAL := 1000.0;                // Y 轴速度上限 [毫米每秒]，域大于 0 / Y axis speed limit
    fNominalCycle : REAL := 0.004;                 // 标称插补周期 [秒]，域 0.0001 到 1 / Nominal interpolation period
    fMaxPathLen   : REAL := 100000.0;              // 允许最大路径长度 [毫米]，域大于 0 / Maximum path length, must exceed zero
END_VAR
VAR_OUTPUT
    bBusy         : BOOL;                          // 插补进行中（含准备段）[-] / Interpolation running, preparation included
    bActive       : BOOL;                          // 位置给定有效（推进中或暂停中）[-] / Position command valid
    bDone         : BOOL;                          // 到达终点，保持到下一次启动 [-] / End reached, held until the next start
    fCmdX         : REAL;                          // X 位置给定 [毫米] / X position command
    fCmdY         : REAL;                          // Y 位置给定 [毫米] / Y position command
    fPathProgress : REAL;                          // 路径完成度 [百分之]，域 0 到 100 / Path progress in percent
    fPathVel      : REAL;                          // 当前合成速度 [毫米每秒] / Current path speed
    fPathLen      : REAL;                          // 本次路径总长 [毫米] / Total path length of this move
    fPeakVel      : REAL;                          // 本次实际峰值速度 [毫米每秒] / Effective peak speed of this move
    bError        : BOOL;                          // 故障级锁存，仅 0204 至 0207 置位 [-] / Latched fault, only fault level codes set it
    uErrorId      : UDINT;                         // 事件码，0 表示无事件 [代码] / Event code, zero means none
    eState        : E_DL_LineInterpPhase;          // 主状态机当前相位 [-] / Current phase of the main state machine
END_VAR
VAR
    fbTrigStart   : R_TRIG;                        // 启动沿检测，主周期无条件刷新 [-] / Start edge detector, refreshed unconditionally
    fbTrigReset   : R_TRIG;                        // 复位沿检测，主周期无条件刷新 [-] / Reset edge detector, refreshed unconditionally
    ePhase        : E_DL_LineInterpPhase := E_DL_LineInterpPhase.eIdle; // 内部相位，对外经 eState 输出 [-] / Internal phase exported as eState
    bInit         : BOOL := FALSE;                 // 首扫标志，初值 FALSE，判据取非 [-] / First-scan flag initialised FALSE
    bFaultLatch   : BOOL;                          // 故障锁存，仅复位分支清除 [-] / Fault latch, cleared by the reset path only
    uErrInt       : UDINT;                         // 故障级码寄存，锁存型 [代码] / Latched fault level code register
    uInfoCode     : UDINT;                         // 本拍信息级码，每拍重算 [代码] / Info level code recomputed every scan
    bDoneLatch    : BOOL;                          // 完成标志保持寄存器 [-] / Done hold register
    fDx           : REAL;                          // X 方向位移 [毫米] / X displacement
    fDy           : REAL;                          // Y 方向位移 [毫米] / Y displacement
    fLen          : REAL;                          // 路径长度 [毫米] / Path length
    fUx           : REAL;                          // X 单位向量分量 [无量纲] / X unit component
    fUy           : REAL;                          // Y 单位向量分量 [无量纲] / Y unit component
    fVEff         : REAL;                          // 生效合成速度 [毫米每秒] / Effective path speed
    fVLimit       : REAL;                          // 单轴限速折算后的合成速度上限 [毫米每秒] / Speed cap derived from axis limits
    fTmpX         : REAL;                          // X 轴限速折算中间量 [毫米每秒] / X cap temporary
    fTmpY         : REAL;                          // Y 轴限速折算中间量 [毫米每秒] / Y cap temporary
    fAccUse       : REAL;                          // 生效加速度 [毫米每二次方秒] / Effective acceleration
    fAccDist      : REAL;                          // 单侧加速距离 [毫米] / One-sided acceleration distance
    fPeak         : REAL;                          // 本次峰值速度 [毫米每秒] / Peak speed of this move
    fVDecelFloor  : REAL;                          // 收尾速度下限 [毫米每秒] / Deceleration speed floor
    fS            : REAL;                          // 当前已走路径位移 [毫米] / Travelled distance
    fV            : REAL;                          // 当前合成速度 [毫米每秒] / Current speed
    fDt           : REAL;                          // 本拍时间增量 [秒] / Time increment of this scan
    bTriangular   : BOOL;                          // 三角曲线标志（无匀速段）[-] / Triangular profile flag
    bNonFinite    : BOOL;                          // 输入含非有限值 [-] / At least one input is not finite
    bSpeedCapped  : BOOL;                          // 单轴限速参与了折算 [-] / An axis limit actually capped the speed
END_VAR
VAR CONSTANT
    DL_LEN_MIN    : REAL := 1.0E-6;                // 判零长度阈值 [毫米] / Zero length threshold
    DL_DT_MIN     : REAL := 1.0E-4;                // 最小插补周期 [秒] / Minimum interpolation period
    DL_DT_MAX     : REAL := 1.0;                   // 最大插补周期 [秒] / Maximum interpolation period
    DL_BIG        : REAL := 1.0E30;                // 非有限判定的大数阈值 [毫米] / Large value threshold for the finiteness test
    DL_DECEL_FLOOR: REAL := 0.05;                  // 收尾速度相对峰值的比例 [无量纲] / Deceleration floor as a fraction of the peak
    DL_PROGRESS_MAX : REAL := 100.0;               // 完成度满值 [百分之] / Full progress value
    DL_TWO        : REAL := 2.0;                   // 实数二，防魔数 [无量纲] / Real two used instead of a magic number
END_VAR

(*------------------------------------------------------------------------------
 * 段 1｜输出确定性默认值（单拍与派生标志每拍预清零，R25 第一律）
 *      Deterministic defaults first, derived flags pre-cleared every scan
 *-----------------------------------------------------------------------------*)
bBusy     := FALSE;                             // 忙碌标志预清零（Busy flag pre-cleared）
bActive   := FALSE;                             // 给定有效标志预清零（Command valid flag pre-cleared）
uInfoCode := 16#0000_0000;                      // 信息级码每拍重算（Info code recomputed every scan）
bNonFinite := FALSE;                            // 非有限标志预清零（Non-finite flag pre-cleared）
bSpeedCapped := FALSE;                          // 限速折算标志预清零（Speed cap flag pre-cleared）

(*------------------------------------------------------------------------------
 * 段 2｜沿检测无条件刷新（红线：实例在 CASE 之外每拍必刷）
 *      Edge detection refreshed unconditionally outside the CASE
 *-----------------------------------------------------------------------------*)
fbTrigStart(CLK := bStart);
fbTrigReset(CLK := bReset);

(*------------------------------------------------------------------------------
 * 段 3｜首扫初始化（唯一合法范式：初值 FALSE，判据取非）
 *      First-scan initialisation following the single legal pattern
 *-----------------------------------------------------------------------------*)
IF NOT bInit THEN
    fS           := 0.0;                        // 位移清零（Travelled distance cleared）
    fV           := 0.0;                        // 速度清零（Speed cleared）
    fUx          := 0.0;                        // X 单位向量清零（X unit component cleared）
    fUy          := 0.0;                        // Y 单位向量清零（Y unit component cleared）
    fLen         := 0.0;                        // 路径长清零（Path length cleared）
    fPeak        := 0.0;                        // 峰值速度清零（Peak speed cleared）
    fAccDist     := 0.0;                        // 加速距离清零（Acceleration distance cleared）
    fAccUse      := DL_TWO;                     // 生效加速度先给安全值（Effective acceleration pre-set to a safe value）
    fDt          := DL_DT_MIN;                  // 时间增量先给下限（Time increment pre-set to the lower bound）
    bTriangular  := FALSE;                      // 三角标志清零（Triangular flag cleared）
    bDoneLatch   := FALSE;                      // 完成保持标志清零（Done hold cleared）
    bFaultLatch  := FALSE;                      // 故障锁存清零（Fault latch cleared）
    uErrInt      := 16#0000_0000;               // 故障码清零（Fault code cleared）
    fPathLen     := 0.0;                        // 路径长出口清零（Path length outlet cleared）
    fPeakVel     := 0.0;                        // 峰值速度出口清零（Peak speed outlet cleared）
    fPathVel     := 0.0;                        // 当前速度出口清零（Current speed outlet cleared）
    fPathProgress:= 0.0;                        // 完成度出口清零（Progress outlet cleared）
    ePhase       := E_DL_LineInterpPhase.eIdle; // 相位复位为待机（Phase reset to idle）
    bInit        := TRUE;                       // 首扫只做一次（First scan runs once）
END_IF

(*------------------------------------------------------------------------------
 * 段 4｜非有限输入前置拦截（NaN 用自身不等于自身判定，无穷用大数阈值判定）
 *      Finiteness gate, NaN by self comparison and infinity by a magnitude bound
 *-----------------------------------------------------------------------------*)
IF (fStartX <> fStartX) OR (fStartY <> fStartY) OR (fEndX <> fEndX) OR (fEndY <> fEndY) THEN
    bNonFinite := TRUE;                         // 坐标含 NaN（A coordinate is NaN）
END_IF
IF (fPathSpeed <> fPathSpeed) OR (fAccel <> fAccel) OR (fMaxSpeedX <> fMaxSpeedX) OR (fMaxSpeedY <> fMaxSpeedY) THEN
    bNonFinite := TRUE;                         // 速度或加速度含 NaN（A speed or acceleration is NaN）
END_IF
IF (ABS(fStartX) > DL_BIG) OR (ABS(fStartY) > DL_BIG) OR (ABS(fEndX) > DL_BIG) OR (ABS(fEndY) > DL_BIG) THEN
    bNonFinite := TRUE;                         // 坐标越出量级上限（A coordinate exceeds the magnitude bound）
END_IF
IF (ABS(fPathSpeed) > DL_BIG) OR (ABS(fAccel) > DL_BIG) OR (ABS(fNominalCycle) > DL_BIG) OR (ABS(fMaxPathLen) > DL_BIG) THEN
    bNonFinite := TRUE;                         // 参数越出量级上限（A parameter exceeds the magnitude bound）
END_IF

(*------------------------------------------------------------------------------
 * 段 5｜标称周期钳位（越界只钳位并置信息级，不停机）
 *      Nominal period clamping with an informational code only
 *-----------------------------------------------------------------------------*)
IF fNominalCycle < DL_DT_MIN THEN
    fDt       := DL_DT_MIN;                     // 周期下限钳位（Clamped to the lower bound）
    uInfoCode := 16#0004_010A;                  // 010A 周期越界已钳位（Period clamped）
ELSIF fNominalCycle > DL_DT_MAX THEN
    fDt       := DL_DT_MAX;                     // 周期上限钳位（Clamped to the upper bound）
    uInfoCode := 16#0004_010A;                  // 010A 周期越界已钳位（Period clamped）
ELSE
    fDt       := fNominalCycle;                 // 合法周期直通（Valid period passed through）
END_IF

(*------------------------------------------------------------------------------
 * 段 6｜使能撤销的最高优先级拦截（先于状态机，切断推进条件）
 *      Enable withdrawal is handled before the state machine
 *-----------------------------------------------------------------------------*)
IF NOT bEnable THEN
    fV := 0.0;                                  // 速度归零（Speed forced to zero）
    IF (ePhase = E_DL_LineInterpPhase.eAccel) OR (ePhase = E_DL_LineInterpPhase.eCruise) OR
       (ePhase = E_DL_LineInterpPhase.eDecel) OR (ePhase = E_DL_LineInterpPhase.eHeld) THEN
        ePhase := E_DL_LineInterpPhase.eIdle;   // 推进中掉使能：回待机（Disabled mid move, back to idle）
        fS     := 0.0;                          // 位移清零，避免下次启动带残留（Distance cleared）
    END_IF
END_IF

(*------------------------------------------------------------------------------
 * 段 7｜主状态机（枚举每个成员均有标签，末尾 ELSE 兜底到终端安全态）
 *      Main state machine, one label per member plus a trailing ELSE fallback
 *-----------------------------------------------------------------------------*)
CASE ePhase OF

    E_DL_LineInterpPhase.eIdle: // 待机：等启动沿，给定停在起点
        fS := 0.0;                              // 位移清零（Distance cleared）
        fV := 0.0;                              // 速度清零（Speed cleared）
        IF bFaultLatch THEN
            ePhase := E_DL_LineInterpPhase.eFault; // 参数已锁故障：进故障态（Gate failed, enter the fault state）
        ELSIF fbTrigStart.Q THEN
            bDoneLatch := FALSE;                // 新一次启动：清完成保持（A new start clears the done hold）
            ePhase     := E_DL_LineInterpPhase.ePrep; // 进准备相（Enter the preparation phase）
        END_IF

    E_DL_LineInterpPhase.ePrep: // 准备：闸门、向量分解、限幅折算、剖面判定
        IF bNonFinite THEN
            IF NOT bFaultLatch THEN
                bFaultLatch := TRUE;            // 锁故障，保留首出码（Latch the fault keeping the first code）
                uErrInt     := 16#0004_0206;    // 0206 输入非有限（Non-finite input）
            END_IF
            bDoneLatch := FALSE;                // 清完成保持（Done hold cleared）
            ePhase     := E_DL_LineInterpPhase.eFault; // 进故障态（Enter the fault state）
        ELSIF (fPathSpeed <= 0.0) OR (fAccel <= 0.0) OR (fMaxSpeedX <= 0.0) OR
              (fMaxSpeedY <= 0.0) OR (fMaxPathLen <= 0.0) THEN
            IF NOT bFaultLatch THEN
                bFaultLatch := TRUE;            // 锁故障（Latch the fault）
                uErrInt     := 16#0004_0204;    // 0204 运动参数非法（Illegal motion parameters）
            END_IF
            bDoneLatch := FALSE;                // 清完成保持（Done hold cleared）
            ePhase     := E_DL_LineInterpPhase.eFault; // 进故障态（Enter the fault state）
        ELSE
            fDx  := fEndX - fStartX;            // X 方向位移（X displacement）
            fDy  := fEndY - fStartY;            // Y 方向位移（Y displacement）
            fLen := SQRT((fDx * fDx) + (fDy * fDy)); // 路径长度（Path length）
            fPathLen := fLen;                   // 路径长出口（Path length outlet）
            IF fLen > fMaxPathLen THEN
                IF NOT bFaultLatch THEN
                    bFaultLatch := TRUE;        // 路径超限：锁故障（Path over the limit, latch a fault）
                    uErrInt     := 16#0004_0205; // 0205 路径超限（Path over the limit）
                END_IF
                bDoneLatch := FALSE;            // 清完成保持（Done hold cleared）
                ePhase     := E_DL_LineInterpPhase.eFault; // 进故障态（Enter the fault state）
            ELSIF fLen < DL_LEN_MIN THEN
                fUx        := 0.0;              // 零长度无单位向量（No unit vector for a zero length move）
                fUy        := 0.0;              // 零长度无单位向量（No unit vector for a zero length move）
                fS         := 0.0;              // 位移为零（No displacement）
                fV         := 0.0;              // 速度为零（No speed）
                fPeak      := 0.0;              // 峰值速度为零（No peak speed）
                bDoneLatch := TRUE;             // 当拍即完成（Completed within this scan）
                uInfoCode  := 16#0004_0109;     // 0109 零长度路径（Zero length path）
                ePhase     := E_DL_LineInterpPhase.eDone; // 直接进完成相（Jump to the done phase）
            ELSE
                fUx := fDx / fLen;              // X 单位向量，除数已过判零闸门（Unit vector, the divisor passed the gate）
                fUy := fDy / fLen;              // Y 单位向量，除数已过判零闸门（Unit vector, the divisor passed the gate）
                fAccUse := fAccel;              // 生效加速度（Effective acceleration）
                fVLimit := fPathSpeed;          // 先与期望合成速度取最小（Start from the desired speed）
                IF ABS(fUx) > DL_LEN_MIN THEN
                    fTmpX := fMaxSpeedX / ABS(fUx); // X 轴折算上限（X cap from the axis limit）
                    IF fTmpX < fVLimit THEN
                        fVLimit      := fTmpX;  // 取更小者（Keep the smaller cap）
                        bSpeedCapped := TRUE;   // 记录限速生效（Record that a cap applied）
                    END_IF
                END_IF
                IF ABS(fUy) > DL_LEN_MIN THEN
                    fTmpY := fMaxSpeedY / ABS(fUy); // Y 轴折算上限（Y cap from the axis limit）
                    IF fTmpY < fVLimit THEN
                        fVLimit      := fTmpY;  // 取更小者（Keep the smaller cap）
                        bSpeedCapped := TRUE;   // 记录限速生效（Record that a cap applied）
                    END_IF
                END_IF
                fVEff     := fVLimit;           // 生效合成速度（Effective path speed）
                fAccDist  := (fVEff * fVEff) / (DL_TWO * fAccUse); // 单侧加速距离（One-sided acceleration distance）
                IF (DL_TWO * fAccDist) > fLen THEN
                    bTriangular := TRUE;        // 两侧之和超过全长：三角曲线（Sum exceeds the path, triangular）
                    fPeak     := SQRT(fAccUse * fLen); // 三角峰值速度（Triangular peak speed）
                    fAccDist  := fLen * 0.5;    // 加速距离取一半（Half of the path）
                    uInfoCode := 16#0004_010C;  // 010C 三角曲线生效（Triangular profile in effect）
                ELSE
                    bTriangular := FALSE;       // 两侧之和不超过全长：梯形曲线（Trapezoidal profile）
                    fPeak       := fVEff;       // 峰值即生效合成速度（Peak equals the effective speed）
                    IF bSpeedCapped THEN
                        uInfoCode := 16#0004_010B; // 010B 单轴限速参与折算（An axis limit capped the speed）
                    END_IF
                END_IF
                fVDecelFloor := fPeak * DL_DECEL_FLOOR; // 收尾速度下限（Deceleration floor）
                fPeakVel     := fPeak;          // 峰值速度出口（Peak speed outlet）
                fS           := 0.0;            // 位移从零起算（Distance starts at zero）
                fV           := 0.0;            // 速度从零起算（Speed starts at zero）
                ePhase       := E_DL_LineInterpPhase.eAccel; // 进加速段（Enter the acceleration segment）
            END_IF
        END_IF

    E_DL_LineInterpPhase.eAccel: // 加速段：速度上升，位移积分
        IF bHold THEN
            fV     := 0.0;                      // 暂停：速度归零（Hold, speed forced to zero）
            ePhase := E_DL_LineInterpPhase.eHeld; // 进暂停相（Enter the held phase）
        ELSE
            fV := MIN(fPeak, fV + (fAccUse * fDt)); // 速度斜坡上升（Ramp the speed up）
            fS := fS + (fV * fDt);              // 位移按速度积分（Integrate the distance）
            (* 出口双条件：位移到加速距离且速度确实升到峰值——暂停恢复后必然满足前者，
               只看位移会当拍跳进匀速段、速度从零直接跳到峰值，故必须同时校验速度 *)
            (* Both conditions are required, otherwise a resume skips the ramp and steps the speed *)
            IF (fS >= fAccDist) AND (fV >= fPeak) THEN
                IF bTriangular THEN
                    ePhase := E_DL_LineInterpPhase.eDecel; // 三角曲线无匀速段（No cruise segment）
                ELSE
                    ePhase := E_DL_LineInterpPhase.eCruise; // 梯形曲线进匀速段（Enter the cruise segment）
                END_IF
            END_IF
        END_IF

    E_DL_LineInterpPhase.eCruise: // 匀速段：速度保持峰值
        IF bHold THEN
            fV     := 0.0;                      // 暂停：速度归零（Hold, speed forced to zero）
            ePhase := E_DL_LineInterpPhase.eHeld; // 进暂停相（Enter the held phase）
        ELSE
            fV := fPeak;                        // 速度保持峰值（Keep the peak speed）
            fS := fS + (fV * fDt);              // 位移按速度积分（Integrate the distance）
            IF fS >= (fLen - fAccDist) THEN
                ePhase := E_DL_LineInterpPhase.eDecel; // 到达减速点（Reach the deceleration point）
            END_IF
        END_IF

    E_DL_LineInterpPhase.eDecel: // 减速段：速度下降到收尾下限，出口钳位到终点
        IF bHold THEN
            fV     := 0.0;                      // 暂停：速度归零（Hold, speed forced to zero）
            ePhase := E_DL_LineInterpPhase.eHeld; // 进暂停相（Enter the held phase）
        ELSE
            fV := MAX(fVDecelFloor, fV - (fAccUse * fDt)); // 速度斜坡下降，保留收尾速度（Ramp down keeping the floor）
            fS := fS + (fV * fDt);              // 位移按速度积分（Integrate the distance）
            IF fS >= fLen THEN
                fS          := fLen;            // 出口钳位，防离散步长超程（Clamp at the end point）
                fV          := 0.0;             // 到位速度归零（Speed zeroed at the end）
                bDoneLatch  := TRUE;            // 完成标志保持（Done hold set）
                fPathProgress := DL_PROGRESS_MAX; // 完成度满值（Progress forced to full）
                ePhase      := E_DL_LineInterpPhase.eDone; // 进完成相（Enter the done phase）
            END_IF
        END_IF

    E_DL_LineInterpPhase.eDone: // 完成：给定等于终点，等下一次启动
        fS          := fLen;                    // 位移停在终点（Distance parked at the end）
        fV          := 0.0;                     // 速度为零（Speed zeroed）
        bDoneLatch  := TRUE;                    // 完成标志保持（Done hold kept）
        fPathProgress := DL_PROGRESS_MAX;       // 完成度满值（Progress full）
        IF fbTrigStart.Q THEN
            bDoneLatch := FALSE;                // 新一次启动：清完成保持（A new start clears the done hold）
            ePhase     := E_DL_LineInterpPhase.ePrep; // 回准备相（Back to preparation）
        END_IF

    E_DL_LineInterpPhase.eHeld: // 暂停：位移保持，恢复后从零速重新加速
        fV := 0.0;                              // 暂停期速度恒为零（Speed stays zero while held）
        IF NOT bHold THEN
            IF (fLen - fS) <= fAccDist THEN
                ePhase := E_DL_LineInterpPhase.eDecel; // 剩余距离已落在减速窗内：直接进减速段，不从零速再加速冲过终点
            ELSE
                ePhase := E_DL_LineInterpPhase.eAccel; // 恢复：从当前位移重新加速（Resume by accelerating from the current distance）
            END_IF
        END_IF

    E_DL_LineInterpPhase.eFault: // 故障：给定保持，等复位沿
        fV := 0.0;                              // 故障期速度为零（Speed zeroed during a fault）

    ELSE
        bFaultLatch := TRUE;                    // 非法状态兜底锁存（Illegal state latched）
        uErrInt     := 16#0004_0207;            // 0207 非法状态兜底（Illegal state fallback code）
        fV          := 0.0;                     // 速度归零（Speed zeroed）
        ePhase      := E_DL_LineInterpPhase.eFault; // 进终端安全态（Enter the terminal safe state）
END_CASE

(*------------------------------------------------------------------------------
 * 段 8｜复位（清故障与完成保持，位移保留供画面诊断）
 *      Reset clears the fault and the done hold, the distance is kept for diagnostics
 *-----------------------------------------------------------------------------*)
IF fbTrigReset.Q THEN
    bFaultLatch := FALSE;                       // 清故障锁存（Clear the fault latch）
    uErrInt     := 16#0000_0000;                // 清故障码（Clear the fault code）
    bDoneLatch  := FALSE;                       // 清完成保持（Clear the done hold）
    fV          := 0.0;                         // 速度归零（Speed zeroed）
    IF (ePhase = E_DL_LineInterpPhase.eFault) THEN
        ePhase := E_DL_LineInterpPhase.eIdle;   // 故障态复位回待机（Fault returns to idle）
        fS     := 0.0;                          // 回待机时位移清零（Distance cleared in idle）
    END_IF
END_IF

(*------------------------------------------------------------------------------
 * 段 9｜给定与派生出口（位置给定按单位向量乘位移，完成度按位移比路径长）
 *      Command and derived outlet mapping
 *-----------------------------------------------------------------------------*)
fCmdX := fStartX + (fUx * fS);                  // X 位置给定（X position command）
fCmdY := fStartY + (fUy * fS);                  // Y 位置给定（Y position command）
IF fLen > DL_LEN_MIN THEN
    fPathProgress := LIMIT(0.0, (fS / fLen) * DL_PROGRESS_MAX, DL_PROGRESS_MAX); // 完成度钳位在 0 到 100（Clamped progress）
ELSIF ePhase = E_DL_LineInterpPhase.eDone THEN
    fPathProgress := DL_PROGRESS_MAX;           // 零长度路径已到达终点：完成度为满值，与完成相口径一致（Zero length already done, full progress）
ELSE
    fPathProgress := 0.0;                       // 其余零长度相位不给百分比，避免除零（No percentage elsewhere, avoids a division by zero）
END_IF
IF (ePhase = E_DL_LineInterpPhase.eAccel) OR (ePhase = E_DL_LineInterpPhase.eCruise) OR (ePhase = E_DL_LineInterpPhase.eDecel) THEN
    bActive   := TRUE;                          // 推进中：给定有效（Moving, the command is valid）
    bBusy     := TRUE;                          // 推进中：忙碌为真（Moving, busy is true）
    fPathVel  := fV;                            // 当前合成速度出口（Current path speed outlet）
ELSIF ePhase = E_DL_LineInterpPhase.eHeld THEN
    bActive   := TRUE;                          // 暂停中：给定仍有效（Held, the command is still valid）
    bBusy     := TRUE;                          // 暂停中：仍算任务未结束（Held, the job is not finished）
    fPathVel  := 0.0;                           // 暂停中合成速度为零（Path speed is zero while held）
ELSIF ePhase = E_DL_LineInterpPhase.ePrep THEN
    bActive   := FALSE;                         // 准备中尚无有效给定（No valid command during preparation）
    bBusy     := TRUE;                          // 准备中算忙碌（Preparation counts as busy）
    fPathVel  := 0.0;                           // 准备中速度为零（Speed is zero during preparation）
ELSE
    bActive   := FALSE;                         // 其余相位无有效给定（No valid command elsewhere）
    fPathVel  := 0.0;                           // 其余相位速度为零（Speed is zero elsewhere）
END_IF
bDone  := bDoneLatch;                           // 完成标志出口（Done outlet）
eState := ePhase;                               // 相位出口（Phase outlet）
bError := bFaultLatch;                          // 故障位只反映故障级锁存（Fault bit reflects the latch only）
IF bError THEN
    uErrorId := uErrInt;                        // 故障级码优先透出（Fault level code has priority）
ELSE
    uErrorId := uInfoCode;                      // 无故障透出本拍信息级码（Info code exposed otherwise）
END_IF
END_FUNCTION_BLOCK

(* ---- FB_DL_MarkPositionLatch.st ---- *)
(*==============================================================================
 * 组件名称 (Component)  : FB_DL_MarkPositionLatch
 * 所属子库 (Sublibrary) : DL_Motion
 * 当前版本 (Version)    : 1.0.0
 * 组件分类 (Category)   : 功能块（FUNCTION_BLOCK）· 标记锁存族 · 色标 / 探针位置锁存
 * 兼容性   (Platform)   : CODESYS 3.5 / TwinCAT 3 / 汇川 InoProShop / Schneider
 *                         Machine Expert；仅依赖 Standard.library
 *                         （R_TRIG / TON / MIN / MAX / ABS），零厂商方言
 * 接口依赖 (Depends)    : I_DL_MotionAxis / E_DL_AxisState（既有契约，Round 05，零修改）
 * 功能描述 (Function)   : 外部标记（色标 / 探针 / 光电开关）触发瞬间锁存轴位置与速度，
 *                         并输出与上次锁存的增量；带布防窗、标记缺失诊断、最近 N 次
 *                         历史环形缓冲。供定长切割、切点相位校正、定长计米与凸轮相位
 *                         补偿前置件使用。
 * 设计要点 (Key notes)  :
 *   ① 位置与速度在同一拍各读一次并同拍锁存，保证两者时间一致（分两拍读会出现
 *      「位置已到、速度还是上一拍」的口径错位）。
 *   ② 本块不累计位置：位置一律来自轴接口，避免与轴侧积分形成双积分漂移。
 *   ③ 一次布防只受理第一条标记沿（连击不重复锁存），去抖交由上游信号处理块承担。
 *   ④ 历史缓冲为定长整体前移写法，用定长 FOR + 深度钳位，不用无界循环。
 *   ⑤ 本块为纯事件型组件：无初始化跟踪语义、无连续量同步逻辑，按库级约定免首扫，
 *      不设首扫标志与跟踪判据（与 FB_DL_SignalDebounce 等事件型件同口径）。
 * 开源溯源 (Origin)     : 原创实现，clean-room。语义来源为 PLCopen 运动控制公开规范中
 *                         的「注册标记 / 探针锁存」工艺概念、公开的色标定长切割与
 *                         追剪技术文章、以及公开的产线节拍链经验总结（来源编号
 *                         RAW_NOTES S-2 相位补偿前置件 / S-14 节拍链）。
 *                         「借鉴对象的许可说明」：上述对象为公开发布但受版权保护的
 *                         规范文档与技术文章，属「可免费查阅、仅借鉴工程语义」类别；
 *                         本实现未复制任何源码，引脚命名、枚举、环形缓冲结构、诊断
 *                         码与状态机 100% 自有设计。
 * 验收向量 (Acceptance) :
 *   V1 布防 → 标记沿 → 锁存位置与速度，首次增量输出为 0；
 *   V2 连续两次布防并触发：第二次增量等于两次锁存位置之差；
 *   V3 布防窗内无标记：超窗进 eMissed，bMarkMissed 为 TRUE（不停机、不置故障）；
 *   V4 重新布防：清 eMissed 与 bMarkMissed，可再次锁存；
 *   V5 nHistoryDepth 填 0：钳位到 1 并出信息级 0170；
 *   V6 清历史：历史缓冲清零，累计标记计数保留；
 *   V7 轴位置为非有限值：锁存 0290，拒绝锁存；
 *   V8 同一布防窗内连击多次：只锁存第一条沿（一次布防一次锁存）。
 * 已知限制 (Limits)     :
 *   ① 布防窗分辨率等于任务扫描周期：窗宽若小于两个扫描周期，实际等效「最多错过
 *      一拍」，属预期行为；极短窗请改用硬件比较输出（探针输入）方案。
 *   ② 本块只用锁存时刻的位置值，不补偿「标记沿到扫描读值」的传输延迟；需要微米
 *      级切点精度时，应由驱动侧探针功能锁存并由本块读取其结果。
 *   ③ 历史缓冲维度以字面量 8 声明（FB 内部常量不能用于其自身引脚声明），运行期
 *      以 UPPER_BOUND / LOWER_BOUND 实测维度做二次钳位。
 * 规格偏离 (Deviation)  :
 *   ① 无（本块引脚与规格逐条一致；未增补任何输入引脚，因纯事件型免首扫）。
 * 红线自检 (Redline)    :
 *   R1 零全局符号区访问 ✓（无全局变量表访问、无外部变量声明）
 *   R2 零物理地址直写 ✓（无输入输出通道地址记号）
 *   R3 纯 IEC 61131-3 ✓（仅 R_TRIG / TON / MIN / MAX / ABS）
 *   R4 防除零 / 防越界 / 浮点容差 ✓（数组索引全程经实测上下界钳位、循环定长、
 *      浮点比较用容差、无除法）
 *   R5 声明行 100% 中英双语同行注释 ✓
 *   R6 ENUM + CASE 且 CASE 含 ELSE 兜底 ✓
 *   R7 边沿与定时器实例无条件周期刷新 ✓（本块无单拍脉冲输出；bLatched /
 *      bMarkMissed 为状态型输出，不跨周期残留）
 *   POU 终结符成对 ✓（FUNCTION_BLOCK ↔ END_FUNCTION_BLOCK，末行即终结符；
 *   TYPE ↔ END_TYPE 成对）
 * 故障码表 (Error codes):
 *   16#0004_0170【信息级】历史深度越界钳位；
 *   16#0004_0171【信息级】布防窗内无标记（缺失提示，与 bMarkMissed 同源）；
 *   16#0004_0290【故障级】轴位置 / 速度非有限值，锁存；
 *   16#0004_0295【故障级】非法状态兜底（本块专用，不与其他块共用）。
 *   信息级码只进 uErrorId；bError 为派生式仅反映 eFault 态。
 * 修订历史 (Revision)   :
 *   2026-11-15  v1.0.0  首版入库（Round 08 · DL_Motion 标记锁存族开族件）
 *============================================================================*)

(*-----------------------------------------------------------------------------
 * 调用示例 (Instance guide)：
 *   fbMark.iAxis := fbConveyorAxis;               // 被采样轴实例注入
 *   fbMark(bEnable := TRUE, tArmWindow := T#5S,
 *          bArm := bCutReady, bTrigger := diColorMark,
 *          nHistoryDepth := 4);
 *   IF fbMark.bLatched THEN
 *       fCutPos := fbMark.fLatchedPos + fCutLength;   // 定长切割：锁存点 + 定长
 *       fCorr   := fbMark.fDeltaPos - fNominalPitch;  // 节距偏差 → 凸轮相位补偿
 *   END_IF
 *   注：标记信号建议先经上游去抖块处理再送入 bTrigger；本块只取上升沿。
 *----------------------------------------------------------------------------*)

(*-----------------------------------------------------------------------------
 * 常见误用与现场提示 (Field notes)：
 *   1 每次切割前都要给一次 bArm 上升沿；不给布防沿则 bTrigger 的沿一律被忽略
 *      （空闲态不收标记），这是「一次布防一次锁存」的刻意语义。
 *   2 布防窗不是「等待时间」而是「超时诊断窗」：窗内没等到标记只提示缺失，
 *      不停机、不置故障，由上层决定是否报警。
 *   3 fDeltaPos 在首个标记时为 0（没有可比对象），不要把它当成「从零点起的位移」；
 *      从零点起的位移请直接读轴位置。
 *   4 累计计数不清零是刻意的：清历史只清位置数组，节拍统计要靠累计计数，
 *      否则换班交接时计数会凭空丢失。
 *   5 轴位置为非有限值时本块直接锁存故障并拒绝锁存，避免把无效值写进历史缓冲
 *      污染后续节距计算。
 *----------------------------------------------------------------------------*)

(*-----------------------------------------------------------------------------
 * 枚举: E_DL_MarkState（归属 DL_Motion，与本功能块同文件发布）
 * 含义: 标记锁存状态机，编号间隔 10 预留扩展位。
 *----------------------------------------------------------------------------*)
{attribute 'strict'}
{attribute 'qualified_only'}
TYPE E_DL_MarkState :
(
    eIdle    := 0,    // 空闲：未布防，忽略触发 / Idle: not armed, triggers ignored
    eArmed   := 10,   // 已布防：等待标记沿 / Armed: waiting for mark edge
    eLatched := 20,   // 已锁存：本周期结果有效，等新布防或复位 / Latched: result valid, waiting for re-arm or reset
    eMissed  := 30,   // 标记缺失：布防窗内无沿（诊断态，非故障） / Missed: no edge within arm window (diagnostic)
    eFault   := 99    // 故障锁存：仅 bReset 上升沿可退出 / Fault: latched, only bReset rising edge exits
) UINT;
END_TYPE

FUNCTION_BLOCK FB_DL_MarkPositionLatch
VAR_INPUT
    bEnable         : BOOL := FALSE;        // 使能（Enable），FALSE=清布防与结果，不影响历史缓冲与累计计数
    bArm            : BOOL := FALSE;        // 布防（Arm），上升沿进入布防态；锁存 / 缺失态下再次上升沿即重新布防
    bTrigger        : BOOL := FALSE;        // 标记输入（Mark input），上升沿为有效标记，电平持续不影响
    tArmWindow      : TIME := T#10S;        // 布防有效窗（Arm window）[ms]，超时未触发转缺失态；T#0S=不限
    bClearHistory   : BOOL := FALSE;        // 清历史缓冲（Clear history），上升沿，不影响累计计数
    bReset          : BOOL := FALSE;        // 复位故障 / 退出缺失态（Reset），上升沿受理
    nHistoryDepth   : UINT := 4;            // 历史深度（History depth）[-]，域 1..实测维度，越界钳位并提示
END_VAR
VAR_OUTPUT
    bLatched        : BOOL := FALSE;        // 已锁存（Latched），仅锁存态为 TRUE
    fLatchedPos     : REAL := 0.0;          // 锁存位置（Latched position）[mm]
    fLatchedSpeed   : REAL := 0.0;          // 锁存瞬间速度（Latched velocity）[mm/s]，带符号
    fDeltaPos       : REAL := 0.0;          // 与上次锁存的位置增量（Delta position）[mm]，无上次时为 0
    bMarkMissed     : BOOL := FALSE;        // 标记缺失（Mark missed），缺失态为 TRUE；重新布防后自动清
    uMarkCount      : UDINT := 0;           // 累计有效标记数（Mark counter）[次]，清历史不影响此计数
    afHistoryPos    : ARRAY[0..7] OF REAL;  // 最近 N 次锁存位置（History positions）[mm]，维度 8，索引 0=最新
    bError          : BOOL := FALSE;        // 故障锁存（Error），派生式仅故障级码参与，信息级码不置位
    uErrorId        : UDINT := 0;           // 故障码（Error code），段位 16#0004_xxxx，0=无故障
END_VAR
VAR_IN_OUT
    iAxis           : I_DL_MotionAxis;      // 被采样轴接口引用（Sampled axis），由调用方注入实现块实例
END_VAR
VAR
    eState          : E_DL_MarkState := E_DL_MarkState.eIdle; // 内部状态机步序（Internal state）
    bFaultLatch     : BOOL := FALSE;        // 故障锁存标志（Fault latch），仅 bReset 沿解除
    bHistValid      : BOOL := FALSE;        // 历史有效标志（History valid），存在可比对的上次锁存
    bWindowOn       : BOOL := FALSE;        // 布防窗计时使能（Arm window timer enable），窗长为 0 时关闭
    bWindowBrk      : BOOL := FALSE;        // 布防窗参数变更标志（Window changed），断输入一拍用
    bIdxOk          : BOOL := FALSE;        // 数组边界有效标志（Index bounds valid），逐拍重算
    fLastPos        : REAL := 0.0;          // 上次锁存位置（Previous latched position）[mm]，增量计算基准
    fPosNow         : REAL := 0.0;          // 本拍轴位置（Axis position this scan）[mm]
    fVelNow         : REAL := 0.0;          // 本拍轴速度（Axis velocity this scan）[mm/s]
    nDepthEff       : DINT := 4;            // 生效历史深度（Effective depth）[-]，已按实测维度钳位
    nLb             : DINT := 0;            // 历史数组下标下界（Array lower bound）[-]，实测取得
    nUb             : DINT := 7;            // 历史数组下标上界（Array upper bound）[-]，实测取得
    nAvail          : DINT := 8;            // 实测可用槽位（Available slots）[-]，上界减下界加一
    nIdx            : DINT := 0;            // 历史搬移索引（Shift index）[-]，循环内使用
    nJ              : DINT := 0;            // 升序循环变量（Ascending loop var，镜像下标用）[-]
    nGuard          : DINT := 0;            // 循环防死锁计数器（Loop guard counter）[-]
    tWindowEff      : TIME := T#10S;        // 生效布防窗（Effective arm window）[ms]，负值归零
    tWindowPrev     : TIME := T#0MS;        // 上拍布防窗（Previous arm window）[ms]，变更检测基准
    fbTrigArm       : R_TRIG;               // 布防指令上升沿（Arm command rising edge）
    fbTrigTrig      : R_TRIG;               // 标记输入上升沿（Mark input rising edge）
    fbTrigClear     : R_TRIG;               // 清历史指令上升沿（Clear history rising edge）
    fbTrigReset     : R_TRIG;               // 复位指令上升沿（Reset command rising edge）
    fbTonArmWindow  : TON;                  // 布防窗超时监控（Arm window timer）
END_VAR
VAR CONSTANT
    DL_MARK_HIST_MAX  : DINT := 8;          // 历史槽位上限（Max history slots）[-]，与引脚声明的字面量维度一致
    DL_MARK_INF_MAX   : REAL := 1.0E30;     // 有限值判定幅值上限（Finite magnitude bound）[无量纲，按比较量量纲同值使用]
    DL_MARK_EPS       : REAL := 1.0E-6;     // 浮点判零容差（Float zero tolerance）[无量纲，按比较量量纲同值使用]
    DL_MARK_DEPTH_MIN : DINT := 1;          // 历史深度下限（Depth lower bound）[-]
    DL_MARK_GUARD_MAX : DINT := 32;         // 循环防死锁上限（Loop guard limit）[-]，远超最大槽位
    DL_MARK_ZERO_TIME : TIME := T#0S;       // 零时间字面量（Zero time literal）[ms]
END_VAR

// 段 1｜边沿与定时器实例无条件周期刷新（红线 R7：严禁置于 IF / CASE 分支内）
fbTrigArm(CLK := bArm);
fbTrigTrig(CLK := bTrigger);
fbTrigClear(CLK := bClearHistory);
fbTrigReset(CLK := bReset);

// 段 2｜出口默认赋值（公约 0.9：早退路径输出必须确定）
bLatched    := FALSE;
bMarkMissed := FALSE;
bError      := (eState = E_DL_MarkState.eFault);

// 段 3｜接口引用有效性防御：未注入轴引用则清输出退出
IF iAxis = 0 THEN
    RETURN;
END_IF

// 段 4｜历史数组实测边界（公约 0.14：数组访问前必须验界）
nLb    := LOWER_BOUND(afHistoryPos, 1);
nUb    := UPPER_BOUND(afHistoryPos, 1);
nAvail := nUb - nLb + 1;
bIdxOk := (nAvail >= DL_MARK_DEPTH_MIN);
IF nAvail > DL_MARK_HIST_MAX THEN
    nAvail := DL_MARK_HIST_MAX;                          // 实测维度超库级上限时按上限钳位，防越界
END_IF

// 段 5｜历史深度钳位（越界钳位并提示，逐拍重算不锁存）
nDepthEff := UINT_TO_DINT(nHistoryDepth);
IF nDepthEff < DL_MARK_DEPTH_MIN THEN
    nDepthEff := DL_MARK_DEPTH_MIN;                      // 低于 1 钳到 1
    uErrorId  := 16#0004_0170;                           // 【信息级】历史深度越界钳位
ELSIF nDepthEff > nAvail THEN
    nDepthEff := nAvail;                                 // 高于实测槽位钳到上界
    uErrorId  := 16#0004_0170;                           // 【信息级】历史深度越界钳位
END_IF

// 段 6｜布防窗参数防御与变更检测（公约 0.6：语义参数变化必须断输入一拍）
IF tArmWindow < DL_MARK_ZERO_TIME THEN
    tWindowEff := DL_MARK_ZERO_TIME;
ELSE
    tWindowEff := tArmWindow;
END_IF
bWindowBrk  := (tWindowEff <> tWindowPrev);              // 窗长变更：本拍断输入，使已计时归零
tWindowPrev := tWindowEff;
bWindowOn   := (tWindowEff > DL_MARK_ZERO_TIME);         // 窗长为 0 表示不限时，不启用计时

// 段 7｜布防窗超时定时器：实例在本行无条件每拍调用（红线 R7），入参先算成普通变量
fbTonArmWindow(IN := (eState = E_DL_MarkState.eArmed) AND bWindowOn AND (NOT bWindowBrk),
               PT := tWindowEff);

// 段 8｜反馈量采集与信号有效性判定
fPosNow := iAxis.fPosition;
fVelNow := iAxis.fVelocity;
IF (fPosNow <> fPosNow) OR (fVelNow <> fVelNow)
   OR (ABS(fPosNow) > DL_MARK_INF_MAX) OR (ABS(fVelNow) > DL_MARK_INF_MAX) THEN
    IF (eState <> E_DL_MarkState.eFault) THEN
        bFaultLatch := TRUE;
        uErrorId    := 16#0004_0290;                     // 【故障级】轴位置 / 速度非有限值
        eState      := E_DL_MarkState.eFault;
    END_IF
END_IF

// 段 9｜使能撤除：清布防与结果（历史缓冲与累计计数保留）
IF NOT bEnable THEN
    eState      := E_DL_MarkState.eIdle;
    bLatched    := FALSE;
    bMarkMissed := FALSE;
END_IF

// 段 10｜清历史沿（只清位置数组，不清累计计数）
IF fbTrigClear.Q AND bIdxOk THEN
    nGuard := 0;
    FOR nIdx := nLb TO nUb DO
        IF nGuard >= DL_MARK_GUARD_MAX THEN
            EXIT;                                        // 防死锁
        END_IF
        nGuard := nGuard + 1;
        afHistoryPos[nIdx] := 0.0;                       // 槽位清零 [mm]
    END_FOR
    bHistValid := FALSE;                                 // 无可比对上次锁存，下次增量输出 0
END_IF

// 段 11｜事件码管理（公约 0.7 / R15）：锁存码仅在解除路径清，瞬时码逐拍重算
IF NOT bFaultLatch THEN
    uErrorId := 0;
END_IF

// 段 12｜主状态机（ENUM + CASE + ELSE 兜底）
CASE eState OF

    E_DL_MarkState.eIdle:                                // 空闲：未布防，忽略标记沿
        bLatched    := FALSE;
        bMarkMissed := FALSE;
        IF fbTrigArm.Q AND bEnable THEN
            bFaultLatch := FALSE;                        // 新布防：锁存码解除路径（R15）
            bMarkMissed := FALSE;
            bLatched    := FALSE;
            eState      := E_DL_MarkState.eArmed;
        ELSIF fbTrigReset.Q THEN
            bFaultLatch := FALSE;
            uErrorId    := 0;
        END_IF

    E_DL_MarkState.eArmed:                               // 已布防：等待标记沿或超窗
        IF fbTrigArm.Q THEN
            bLatched := FALSE;                           // 重复布防：重新计时（一次布防一次锁存）
        ELSIF fbTrigTrig.Q THEN
            // 同一拍各读一次位置与速度，保证同拍一致
            fLatchedPos   := fPosNow;                    // 锁存位置 [mm]
            fLatchedSpeed := fVelNow;                    // 锁存速度 [mm/s]
            IF bHistValid THEN
                fDeltaPos := fLatchedPos - fLastPos;     // 与上次锁存的增量 [mm]
            ELSE
                fDeltaPos := 0.0;                        // 首个标记无对比对象，增量输出 0
            END_IF
            fLastPos   := fLatchedPos;                   // 增量基准推进 [mm]
            bHistValid := TRUE;
            // 历史缓冲头插（整体前移，定长循环 + 实测边界）
            IF bIdxOk AND (nDepthEff >= DL_MARK_DEPTH_MIN) THEN
                nGuard := 0;
                FOR nJ := DL_MARK_DEPTH_MIN TO (nDepthEff - 1) DO
                    nIdx := (nDepthEff - 1) - nJ + DL_MARK_DEPTH_MIN;   // 镜像下标：R509 禁 DOWNTO（Mirrored index, DOWNTO unsupported）
                    IF nGuard >= DL_MARK_GUARD_MAX THEN
                        EXIT;                            // 防死锁
                    END_IF
                    nGuard := nGuard + 1;
                    IF (nLb + nIdx) <= nUb THEN
                        afHistoryPos[nLb + nIdx] := afHistoryPos[nLb + nIdx - 1]; // 槽位后移
                    END_IF
                END_FOR
                afHistoryPos[nLb] := fLatchedPos;        // 最新值写入 0 号槽 [mm]
            END_IF
            IF uMarkCount < 16#FFFF_FFFF THEN
                uMarkCount := uMarkCount + 1;            // 累计有效标记数 [次]，饱和不加
            END_IF
            bLatched := TRUE;
            eState   := E_DL_MarkState.eLatched;
        ELSIF fbTonArmWindow.Q THEN
            bMarkMissed := TRUE;                         // 超窗无标记：诊断态，停机与否由上层决定
            uErrorId    := 16#0004_0171;                 // 【信息级】布防窗内无标记
            eState      := E_DL_MarkState.eMissed;
        END_IF

    E_DL_MarkState.eLatched:                             // 已锁存：结果保持，等新布防或复位
        bLatched := TRUE;
        IF fbTrigArm.Q AND bEnable THEN
            bLatched := FALSE;
            eState   := E_DL_MarkState.eArmed;           // 重新布防
        ELSIF fbTrigReset.Q THEN
            bLatched := FALSE;
            eState   := E_DL_MarkState.eIdle;
        END_IF

    E_DL_MarkState.eMissed:                              // 标记缺失：等重新布防或复位
        bMarkMissed := TRUE;
        IF fbTrigArm.Q AND bEnable THEN
            bMarkMissed := FALSE;
            bLatched    := FALSE;
            eState      := E_DL_MarkState.eArmed;        // 重新布防即清缺失
        ELSIF fbTrigReset.Q THEN
            bMarkMissed := FALSE;
            uErrorId    := 0;
            eState      := E_DL_MarkState.eIdle;
        END_IF

    E_DL_MarkState.eFault:                               // 故障锁存：仅复位沿可退出
        bLatched    := FALSE;
        bMarkMissed := FALSE;
        IF fbTrigReset.Q THEN
            bFaultLatch := FALSE;                        // 唯一解除路径
            uErrorId    := 0;
            eState      := E_DL_MarkState.eIdle;
        END_IF

    ELSE                                                 // 非法状态兜底（本块专用码）
        bFaultLatch := TRUE;
        uErrorId    := 16#0004_0295;                     // 【故障级】非法状态兜底
        bLatched    := FALSE;
        bMarkMissed := FALSE;
        eState      := E_DL_MarkState.eFault;

END_CASE

// 段 13｜出口映射（派生式，信息级码不参与 bError）
bError      := (eState = E_DL_MarkState.eFault);
bLatched    := (eState = E_DL_MarkState.eLatched);
bMarkMissed := (eState = E_DL_MarkState.eMissed);

END_FUNCTION_BLOCK

(* ---- FB_DL_MeasureInputLatch.st ---- *)
(*==============================================================================
 * 组件名称 (Component)  : FB_DL_MeasureInputLatch
 * 所属子库 (Sublibrary) : DL_Motion ｜ 版本 (Version) : 1.0.0 ｜ 2026-11-24
 * 码位     (Code Segment): 16#0005_21C0（DL_Motion 段内 21xx 子带）
 * 复杂度   (Complexity) : C3
 * 兼容性   (Platform)   : CODESYS 3.5+ / TwinCAT 3 / 汇川 InoProShop / 施耐德 Machine Expert
 *                         仅依赖 IEC 61131-3 标准库（TON / R_TRIG / ABS / REAL_TO_LREAL /
 *                         LREAL_TO_REAL），零厂商私有库
 * 开源溯源 (Provenance) : ThorstenBrach/SRCI_CLIENT_PLC / MC_MeasuringInputFB / MIT /
 *                         借鉴点：测量输入「布防—触发—锁存—读取」的相序与布防窗口超时语义
 *                         （未复制任何实现行，按 IEC 61131-3 重写为五相状态机 + 软件边沿锁存）
 * 功能描述 (Function)   : 探针测量输入锁存。收到布防命令（bArm 上升沿）后进入 eArmed，等探针原始
 *                         信号上升沿：若该沿落在有效窗口 [rWindowStartMm, rWindowEndMm] 内，
 *                         把当时的 rAxisPosMm 锁存为 rLatchPosMm 并置 bLatched；窗口外触发只
 *                         累加 iOutsideCnt 并继续等待（不清布防，避免一个毛刺废掉整次测量）。
 *                         锁存后经 tLatchHold 保持相把结果留在出口供上层读取，然后自动解除布防
 *                         回 eIdle，等下一轮 bArm 沿。
 *                         **边沿纪律（R79 教训）**：bArm 与 bProbeRaw 一律 R_TRIG 取上升沿。
 *                         电平布防会在同一 bArm 电平内反复重新布防，把后续毛刺重复锁存；电平
 *                         探针同理。两者都在 CASE 外无条件刷新（R7），CASE 内只读 .Q。
 *                         **布防超时兜底（R448/R449）**：eArmed 是唯一的外部事件等待相，若一直
 *                         无触发则相驻留无界，故用 tonArm（PT := tArmTimeout）兜底 → 故障级 51。
 *                         **bEnable = FALSE 语义（R191 二选一，本件选「降级为安全值 + 置标志」）**：
 *                         布防与锁存位撤销、bDone 归假、相位回 eIdle；rLatchPosMm 与两计数保留
 *                         （已发生的测量事实不撤回，仅由 bReset 沿清计数器）。
 * 接口     (Interface)  : 输入 bEnable / bReset（上升沿）/ bArm（上升沿有效）/ bProbeRaw（上升沿
 *                         有效）/ rAxisPosMm / rWindowStartMm / rWindowEndMm / tArmTimeout /
 *                         tLatchHold；输出 eState（E_DL_MeasureInputLatch_State）/ bArmed /
 *                         bLatched / bDone（锁存单拍）/ bError / iErrCode / rLatchPosMm /
 *                         iOutsideCnt / iEdgeCnt。
 * 状态迁移表 (State Transition Table)：
 *   ① eIdle → eArmed：bEnable 且 rtArm.Q（布防上升沿）且窗口合法且无锁存；拍 N 进入 /
 *      本拍行为：拒绝锁存与完成位，保留上次 rLatchPosMm 供读取 / 拍 N+1 转出至 eArmed。
 *   ② eArmed → eArmed（驻留）：rtProbe.Q 且该沿落在窗口外；拍 N 进入 / 本拍行为：iEdgeCnt+1、
 *      iOutsideCnt+1，拒绝锁存（毛刺不废测量）/ 拍 N+1 驻留继续等待。
 *   ③ eArmed → eLatched：rtProbe.Q 且 rAxisPosMm 落在 [窗口起点 − 容差, 窗口终点 + 容差]；
 *      拍 N 进入 / 本拍行为：iEdgeCnt+1、rLatchPosMm 写入本拍轴位置（本拍合法事件优先于超时，
 *      R275）/ 拍 N+1 转出至 eLatched。
 *   ④ eArmed → eIdle：bEnable = FALSE（进相前置条件消失，第二出口，R98）。
 *   ⑤ eArmed → eFault：tonArm.Q（布防窗口内无触发，故障级 51）。
 *   ⑥ eLatched → eHold：单拍置位；拍 N 进入 / 本拍行为：bLatched 与 bDone 置单拍、布防解除、
 *      拒收新沿 / 拍 N+1 转出至 eHold。
 *   ⑦ eHold → eIdle：tonHold.Q（保持到期，自动解除布防）；拍 N 进入 / 本拍行为：bLatched 归假、
 *      拒绝新锁存（须重新布防）/ 拍 N+1 转出至 eIdle。
 *   ⑧ eHold → eIdle：bEnable = FALSE（第二出口）。
 *   ⑨ 任意相 → eFault：窗口参数非法或非有限（52）；轴位置非有限（53）；非法枚举（99）。
 *      锁存后由段 7 段尾迁移闸迁相。
 *   ⑩ eFault → eIdle：bReset 上升沿；拍 N 进入 / 本拍行为：清锁存、错误码、布防与锁存位与
 *      两计数，**保留** rLatchPosMm / 拍 N+1 转出至 eIdle。出口穷举、不滞留故障态。
 * 边界     (Boundary)   : ① 两个 TON 与两个 R_TRIG 全部在 CASE 外无条件调用（R7）；TON 的 IN 均含
 *                            NOT .Q 自复位项（R188），禁靠外部沿清零。
 *                         ② 同拍双窗配比约束（R100）：tonArm（PT := _tArm）覆盖 eArmed 相，
 *                            tonHold（PT := _tHold）覆盖 eHold 相，两使能域互斥不相交，无竞态；
 *                            配置建议 tLatchHold ≤ tArmTimeout（读取保持不得长于布防等待，
 *                            否则上层会同时看到上一轮保持与本轮布防）。
 *                         ③ 组态域闸全覆盖（FB51-2）：三个浮点入参 rAxisPosMm / rWindowStartMm /
 *                            rWindowEndMm 全部逐项枚举；非有限判定用自反 x <> x 与差值自减
 *                            (x−x) <> (x−x) 双判，禁用近似阈值与 ABS(x−x) 形态（R4 / R79）。
 *                         ④ 窗口判据带容差：下沿 `_fPos >= (_fWinStart - 1.0E-6)`、上沿
 *                            `_fPos <= (_fWinEnd + 1.0E-6)`，禁 `=` / `<>` 判等（R4）。
 *                         ⑤ 窗口合法性闸（终点 > 起点）与轴位置非有限闸在整个运行期每拍生效，
 *                            不只在布防拍判定——运行中把窗口改反同样立即锁存（域闸不偷工）。
 *                         ⑥ 时间参数两级回退（FB32-3）：越域回默认常量（各自在有效域内），
 *                            故无需二级钳定；回退不置故障（不新增码位）。
 *                         ⑦ 零全局耦合（无 GVL / VAR_EXTERNAL / %I / %Q，R1 / R2）。
 * 码表     (Codes)      : 本件按派单指定使用小整数码。信息级（永不置 bError）：无。
 *                         故障级（置 bError，锁存至 bReset 沿）：
 *                         51 = 布防窗口内无触发超时；反证：该场景下 bArmed 恒真、bLatched 恒假、
 *                              两计数不变，与「正在等探针」的输出组合完全同形，只能靠码区分。
 *                         52 = 窗口参数非法（终点 ≤ 起点，或窗口端点非有限）；反证：该场景
 *                              窗口判据退化为空集或全域，锁存位行为与「探针一直不来」同形，
 *                              且补救动作是改参数而非查探针，必须独立成码。
 *                         53 = 轴位置非有限（编码器失效或位置回读断链）；反证：与 52 的区别是
 *                              参数正确而回读崩塌，补救动作是查反馈而非改参数，须独立成码。
 *                         99 = 非法状态枚举值（ELSE 兜底）。
 * 分工声明 (Scope)      : 轴的实际位置回读与编码器健康监测归 DL_Motion 轴类件（本件只消费
 *                         rAxisPosMm）；探针硬件滤波（去抖 / 脉宽门限）归输入模块组态或硬件
 *                         滤波层（本件只做软件上升沿与窗口裁决）；采点数据的工艺解释与补偿
 *                         计算归上层测量应用件。本件只做**一次测量的布防—锁存—读取时序**。
 * 归属     (Ownership)  : E_DL_MeasureInputLatch_State 归属本文件（全库唯一定义，R264）。
 * 命名偏离 (Naming Ex.) : 本件按派单原文保留 r 前缀表示 REAL（rAxisPosMm / rWindowStartMm /
 *                         rWindowEndMm / rLatchPosMm），i 前缀表示 INT（iErrCode / iOutsideCnt /
 *                         iEdgeCnt）；内部计算升位为 LREAL 的 f 前缀。与规范 1.2 节 n 前缀存在
 *                         登记偏离，接口契约优先不改名。
 * 红线自检 (Redline)    : R1 ✓ 零 GVL / VAR_EXTERNAL ｜ R2 ✓ 零 %I/%Q（探针为普通引脚，非物理
 *                         地址）｜ R3 ✓ 纯 IEC 61131-3（TON / R_TRIG / ABS / REAL_TO_LREAL /
 *                         LREAL_TO_REAL）｜ R4 ✓ 无除法 + 窗口判据带容差 + 自反/差值双判非有限
 *                         ｜ R5 ✓ 逐行同行中英双语注释 ｜ R6 ✓ 五态 ENUM + CASE + ELSE 兜底
 *                         ｜ R7 ✓ TON / R_TRIG 全在 CASE 外无条件调用 ｜ R8 ✓ 无 METHOD（全内联）
 *                         ｜ R10 ✓ 无构造式转换（仅标准转换函数）｜ R11 ✓ 声明全分号结尾
 *                         ｜ R12 ✓ ENUM 成员用 := ｜ R14 ✓ 无 PROPERTY ｜ R16 ✓ 不引用任何外部 FB/FC。
 * 修订历史 (Revision)   : 2026-11-24  v1.0.0  R81-B 首版
 * 验收向量 (Acceptance) :
 *   V1 窗口内正常锁存：rWindowStartMm=10.0、rWindowEndMm=20.0、tArmTimeout=T#2S、
 *      tLatchHold=T#200MS；bEnable=TRUE 后 bArm 起一沿 → eState=eArmed、bArmed=TRUE；
 *      轴到 15.0 时探针起沿 → rLatchPosMm=15.0、bLatched=TRUE、bDone 单拍、iEdgeCnt=1、
 *      iOutsideCnt=0；保持 200ms 后 eState=eIdle、bArmed=FALSE、bLatched=FALSE。
 *   V2 窗口外触发不废测量：轴到 5.0 时探针起沿 → iEdgeCnt=1、iOutsideCnt=1、eState 仍 eArmed、
 *      bLatched=FALSE；随后轴到 18.0 再起沿 → rLatchPosMm=18.0、iEdgeCnt=2、iOutsideCnt=1。
 *   V3 布防超时：bArm 起沿后探针永不来、tArmTimeout=T#1S → 1s 后 eState=eFault、iErrCode=51、
 *      bError=TRUE、bArmed=FALSE；bReset 上升沿 → eState=eIdle、bError=FALSE、iEdgeCnt 归零、
 *      rLatchPosMm 保持 18.0（不清）。
 *   V4 窗口倒置：rWindowStartMm=20.0、rWindowEndMm=10.0 → eState=eFault、iErrCode=52、
 *      bError=TRUE（无需等布防沿，运行期每拍生效）。
 *   V5 边沿纪律：bArm 保持 TRUE 电平不动、探针抖动三次 → 只锁存第一次有效沿（iEdgeCnt 按实际
 *      上升沿计），bDone 仅一拍；撤 bArm 再起才进入下一轮。
 *   V6 撤使能：eArmed 中 bEnable=FALSE → eState=eIdle、bArmed=FALSE、bError=FALSE、
 *      iEdgeCnt / iOutsideCnt 保持。
 *============================================================================*)

(*-----------------------------------------------------------------------------
 * 枚举: E_DL_MeasureInputLatch_State（探针测量输入锁存相位；eFault 为安全相）
 *----------------------------------------------------------------------------*)
TYPE E_DL_MeasureInputLatch_State :
(
    eIdle   := 0,     // 空闲：等布防命令上升沿 / Idle: waiting for the arm command rising edge
    eArmed  := 10,    // 布防相：等探针上升沿，窗口内锁存、窗口外继续等 / Armed: waiting for the probe edge, latch inside the window
    eLatched := 20,   // 锁存相：单拍置锁存与完成 / Latched: one-scan latch and completion
    eHold   := 30,    // 保持相：把结果留在出口，到期自动解除布防 / Hold: keeping the result readable until the hold expires
    eFault  := 90     // 故障安全相：锁存成因，布防与锁存全撤 / Fault safe phase: latched cause, arm and latch withdrawn
);
END_TYPE

FUNCTION_BLOCK FB_DL_MeasureInputLatch
VAR_INPUT
    bEnable       : BOOL := FALSE;      // 使能：FALSE 撤销布防与锁存并回空闲 / Enable, FALSE withdraws arm and latch and returns to idle
    bReset        : BOOL := FALSE;      // 复位（上升沿；清锁存/布防/两计数，不清上次锁存位置）/ Reset rising edge clearing latch, arm and counters but not the last latched position
    bArm          : BOOL := FALSE;      // 布防命令（上升沿有效）/ Arm command, rising edge only
    bProbeRaw     : BOOL := FALSE;      // 探针原始信号（上升沿有效）/ Raw probe signal, rising edge only
    rAxisPosMm    : REAL := 0.0;        // 轴当前位置回读 [mm] / Current axis position feedback
    rWindowStartMm : REAL := 0.0;       // 有效窗口起点，须 < 终点 [mm] / Valid window start, strictly below the end
    rWindowEndMm  : REAL := 100.0;      // 有效窗口终点，须 > 起点 [mm] / Valid window end, strictly above the start
    tArmTimeout   : TIME := T#5S;       // 布防等待上限，有效域 10ms..10min [s] / Arming wait limit, valid domain 10 ms through 10 min
    tLatchHold    : TIME := T#200MS;    // 锁存结果保持时长，有效域 10ms..10min [s] / Latch hold duration, valid domain 10 ms through 10 min
END_VAR
VAR_OUTPUT
    eState        : E_DL_MeasureInputLatch_State;   // 当前相位出口（段 8 单点映射）/ Current phase outlet mapped once at segment 8
    bArmed        : BOOL;               // 布防中（仅 eArmed 相为真）/ Armed, true only inside the eArmed phase
    bLatched      : BOOL;               // 锁存有效（eLatched 起至保持到期）/ Latch valid from eLatched until the hold expires
    bDone         : BOOL;               // 锁存完成单拍脉冲 / One-scan latch completion pulse
    bError        : BOOL;               // 故障锁存标志 / Fault latch flag
    iErrCode      : INT := 0;           // 错误码（故障期锁存回放，其余拍为 0）/ Error code, latched code replayed while in fault
    rLatchPosMm   : REAL := 0.0;        // 锁存位置（保留至下一次锁存，复位不清）[mm] / Latched position kept until the next latch and across resets
    iOutsideCnt   : INT := 0;           // 窗口外触发累计 [次] / Cumulative out-of-window trigger count
    iEdgeCnt      : INT := 0;           // 探针上升沿累计（含窗口外）[次] / Cumulative probe rising edges including out-of-window ones
END_VAR
VAR
    _eState       : E_DL_MeasureInputLatch_State := E_DL_MeasureInputLatch_State.eIdle;   // 内部相位（CASE 唯一写入目标）/ Internal phase, the only CASE write target
    _bFaultLatch  : BOOL := FALSE;      // 故障锁存位（仅 bReset 上升沿清除）/ Fault latch bit, cleared only by the bReset rising edge
    _iErrLatch    : INT := 0;           // 锁存故障码（故障期唯一回放源，FB33-1）/ Latched fault code, the only replay source during fault
    _iErrTmp      : INT := 0;           // 当拍故障首因中间量 / First fault cause of this scan
    _bFaultReq    : BOOL := FALSE;      // 当拍故障请求标志（段 7 统一锁存）/ Fault request of this scan latched at segment 7
    _bCfgOk       : BOOL := TRUE;       // 窗口与位置闸通过标志 / Window and position gate flag
    _bLatchedLatch : BOOL := FALSE;     // 锁存保持量（eLatched 置位，eHold 到期清）/ Latch holding bit set in eLatched and cleared when the hold expires
    _bDonePulse   : BOOL := FALSE;      // 完成内部单拍位（段 1 预置，段 8 映射）/ Internal one-scan done bit preset at segment 1
    _fPos         : LREAL := 0.0;       // 轴位置升位副本 [mm] / Promoted copy of the axis position
    _fWinStart    : LREAL := 0.0;       // 窗口起点升位副本 [mm] / Promoted copy of the window start
    _fWinEnd      : LREAL := 0.0;       // 窗口终点升位副本 [mm] / Promoted copy of the window end
    _fLatchPos    : LREAL := 0.0;       // 锁存位置保持量（升位）[mm] / Holding value of the latched position, promoted
    _iOutsideCnt  : INT := 0;           // 内部窗口外触发累计 [次] / Internal out-of-window trigger counter
    _iEdgeCnt     : INT := 0;           // 内部探针上升沿累计 [次] / Internal probe rising-edge counter
    _tArm         : TIME := T#5S;       // 布防等待上限钳定值（两级回退结果）[s] / Clamped arming limit after the two-level fallback
    _tHold        : TIME := T#200MS;    // 保持时长钳定值（两级回退结果）[s] / Clamped hold duration after the two-level fallback
    rtReset       : R_TRIG;             // bReset 边沿实例（段 5 无条件调用，R18）/ bReset edge instance called unconditionally
    rtArm         : R_TRIG;             // 布防命令边沿实例（段 5 无条件调用，防电平重复布防，R79）/ Arm edge instance preventing level re-arming
    rtProbe       : R_TRIG;             // 探针边沿实例（段 5 无条件调用，防毛刺电平抖动）/ Probe edge instance suppressing level chatter
    tonArm        : TON;                // 布防等待超时计时器（段 5 无条件调用）/ Arming timeout timer called unconditionally
    tonHold       : TON;                // 锁存结果保持计时器（段 5 无条件调用）/ Latch hold timer called unconditionally
END_VAR
VAR CONSTANT
    DL_MIL_ZERO      : LREAL := 0.0;                // 浮点零基准（作有限性判据的对照量）[-] / Float zero used as the finiteness reference
    DL_MIL_EPS       : LREAL := 1.0E-6;             // 位置比较容差，微米级 [mm] / Position comparison tolerance at the micrometre level
    DL_MIL_T_MIN     : TIME := T#10MS;              // 时间参数下限 [s] / Time parameter lower bound
    DL_MIL_T_MAX     : TIME := T#10M;               // 时间参数上限 [s] / Time parameter upper bound
    DL_MIL_ARM_DEF   : TIME := T#5S;                // 布防等待上限默认回退值（本身在域内）[s] / Default fallback arming limit, already inside the domain
    DL_MIL_HOLD_DEF  : TIME := T#200MS;             // 保持时长默认回退值（本身在域内）[s] / Default fallback hold duration, already inside the domain
    DL_MIL_ONE       : INT := 1;                    // 计数步进一 [次] / Counter step of one
END_VAR

(* —— 段 1：中间量预置（只清单拍标志与扫描量，不清锁存位 / 保持位置 / 两计数，FB32-1） —— *)
_iErrTmp    := 0;                          // 当拍故障首因复位 / Scan first fault cause reset
_bFaultReq  := FALSE;                      // 当拍故障请求复位 / Scan fault request reset
_bCfgOk     := TRUE;                       // 闸标志复位 / Gate flag reset
_bDonePulse := FALSE;                      // 完成单拍位预置（单拍路径唯一预置点，FB51-8）/ Done pulse preset, the single preset point

(* —— 段 2：REAL 入参升位（R10 标准转换，内部一律 LREAL 运算） —— *)
_fPos      := REAL_TO_LREAL(rAxisPosMm);        // 位置升位 / Position promoted
_fWinStart := REAL_TO_LREAL(rWindowStartMm);    // 窗口起点升位 / Window start promoted
_fWinEnd   := REAL_TO_LREAL(rWindowEndMm);      // 窗口终点升位 / Window end promoted

(* —— 段 3：时间参数两级回退（越域回默认常量，默认常量在域内故无需二级钳定，FB32-3） —— *)
IF (tArmTimeout < DL_MIL_T_MIN) OR (tArmTimeout > DL_MIL_T_MAX) THEN
    _tArm := DL_MIL_ARM_DEF;               // 越域：回一级默认常量 / Out of domain: fall back to the default constant
ELSE
    _tArm := tArmTimeout;                  // 域内：原值采用 / Inside the domain: take the value as given
END_IF
IF (tLatchHold < DL_MIL_T_MIN) OR (tLatchHold > DL_MIL_T_MAX) THEN
    _tHold := DL_MIL_HOLD_DEF;             // 越域：回一级默认常量 / Out of domain: fall back to the default constant
ELSE
    _tHold := tLatchHold;                  // 域内：原值采用 / Inside the domain: take the value as given
END_IF

(* —— 段 4：组态域闸全覆盖（三个浮点入参逐项枚举，FB51-2；非有限双判，R4 / R79） —— *)
IF (_fWinStart <> _fWinStart) OR ((_fWinStart - _fWinStart) <> (_fWinStart - _fWinStart)) THEN
    _bCfgOk  := FALSE;                     // 窗口起点非有限 / Window start is not finite
    _iErrTmp := 52;                        // 故障级：窗口参数非法 / Fault: illegal window parameter
END_IF
IF _bCfgOk THEN
    IF (_fWinEnd <> _fWinEnd) OR ((_fWinEnd - _fWinEnd) <> (_fWinEnd - _fWinEnd)) THEN
        _bCfgOk  := FALSE;                 // 窗口终点非有限 / Window end is not finite
        _iErrTmp := 52;                    // 故障级：窗口参数非法 / Fault: illegal window parameter
    END_IF
END_IF
IF _bCfgOk THEN
    IF (_fWinEnd - _fWinStart) <= DL_MIL_EPS THEN
        _bCfgOk  := FALSE;                 // 窗口倒置或退化（终点须严格大于起点）/ Inverted or degenerate window, the end must exceed the start
        _iErrTmp := 52;                    // 故障级：窗口参数非法 / Fault: illegal window parameter
    END_IF
END_IF
IF _bCfgOk THEN
    IF (_fPos <> _fPos) OR ((_fPos - _fPos) <> (_fPos - _fPos)) THEN
        _bCfgOk  := FALSE;                 // 轴位置非有限（编码器失效）/ Axis position is not finite
        _iErrTmp := 53;                    // 故障级：轴位置非有限 / Fault: non-finite axis position
    END_IF
END_IF

(* —— 段 5：边沿与定时器（CASE 外无条件调用，R7；TON 的 IN 含 NOT .Q 自复位，R188） —— *)
rtReset(CLK := bReset);                    // bReset 边沿无条件刷新（R18）/ bReset edge refreshed unconditionally
rtArm(CLK := bArm);                        // 布防命令边沿无条件刷新（防电平重复布防，R79）/ Arm edge refreshed unconditionally
rtProbe(CLK := bProbeRaw);                 // 探针边沿无条件刷新（防电平抖动重复计数）/ Probe edge refreshed unconditionally
tonArm(IN := (_eState = E_DL_MeasureInputLatch_State.eArmed) AND (NOT tonArm.Q) AND (NOT _bFaultLatch),
       PT := _tArm);                       // 布防等待超时（自复位后逐轮再起）/ Arming timeout retriggered each round
tonHold(IN := (_eState = E_DL_MeasureInputLatch_State.eHold) AND (NOT tonHold.Q) AND (NOT _bFaultLatch),
        PT := _tHold);                     // 锁存结果保持计时 / Latch hold timer

(* —— 段 6：状态机主体（唯一相位写入点；故障只置请求，锁存与迁相由段 7 执行，R21） —— *)
CASE _eState OF
    E_DL_MeasureInputLatch_State.eIdle :
        (* 迁移①：布防沿 + 窗口与位置闸通过 → 布防相；保留上次锁存位置供上层读取 *)
        IF bEnable AND rtArm.Q AND _bCfgOk AND (NOT _bFaultLatch) THEN
            _eState := E_DL_MeasureInputLatch_State.eArmed;        // 进布防相 / Move to the armed phase
        END_IF

    E_DL_MeasureInputLatch_State.eArmed :
        (* 同拍竞态处理：本拍探针沿优先于超时迁移（R275），超时判定列最后 *)
        IF rtProbe.Q THEN
            _iEdgeCnt := _iEdgeCnt + DL_MIL_ONE;                   // 沿计数（含窗口外）/ Edge counted including out-of-window events
            IF (_fPos >= (_fWinStart - DL_MIL_EPS)) AND (_fPos <= (_fWinEnd + DL_MIL_EPS)) THEN
                _fLatchPos := _fPos;                               // 窗口内：锁存本拍轴位置（唯一写入点）/ Inside the window: latch the position, the single write point
                _eState    := E_DL_MeasureInputLatch_State.eLatched;   // 迁移③：进锁存相 / Move to latched
            ELSE
                _iOutsideCnt := _iOutsideCnt + DL_MIL_ONE;          // 窗口外：只计数，继续等待（毛刺不废测量）/ Out of window: count only and keep waiting
            END_IF
        ELSIF tonArm.Q THEN
            _iErrTmp   := 51;                                      // 故障级：布防窗口内无触发 / Fault: no trigger inside the arming window
            _bFaultReq := TRUE;                                    // 请求段 7 锁存 / Request the latch at segment 7
        ELSIF NOT bEnable THEN
            _eState := E_DL_MeasureInputLatch_State.eIdle;          // 迁移④：前置条件消失回空闲 / Precondition gone, back to idle
        END_IF

    E_DL_MeasureInputLatch_State.eLatched :
        (* 迁移⑥：单拍置位；拍 N 进入 / 本拍行为：bLatched 与 bDone 各置一次、布防解除 / 拍 N+1 转出至 eHold *)
        _bLatchedLatch := TRUE;                                        // 锁存保持量置位（段 8 映射）/ Latch holding bit raised and mapped at segment 8
        _bDonePulse    := TRUE;                                        // 完成内部单拍置位（段 8 映射）/ Internal done pulse raised and mapped at segment 8
        _eState        := E_DL_MeasureInputLatch_State.eHold;           // 迁移⑥：进保持相 / Move to hold

    E_DL_MeasureInputLatch_State.eHold :
        (* 迁移⑦/⑧：保持到期自动解除布防，或失能立即解除 *)
        IF tonHold.Q THEN
            _bLatchedLatch := FALSE;                                   // 保持到期：锁存位归假（须重新布防）/ Hold expired: latch cleared, re-arming required
            _eState        := E_DL_MeasureInputLatch_State.eIdle;       // 迁移⑦：回空闲相 / Back to idle
        ELSIF NOT bEnable THEN
            _bLatchedLatch := FALSE;                                   // 失能：锁存位归假 / Disabled: latch cleared
            _eState        := E_DL_MeasureInputLatch_State.eIdle;       // 迁移⑧：回空闲相 / Back to idle
        END_IF

    E_DL_MeasureInputLatch_State.eFault :
        (* 迁移⑩：复位沿出口（唯一出口，穷举可达）；锁存位置保留
           拍 N 进入 / 本拍行为：清锁存、错误码、布防位与两计数 / 拍 N+1 转出至 eIdle *)
        IF rtReset.Q THEN
            _bFaultLatch   := FALSE;                                   // 清故障锁存 / Clear the fault latch
            _iErrLatch     := 0;                                       // 清锁存故障码 / Clear the latched fault code
            _bLatchedLatch := FALSE;                                   // 清锁存保持量 / Clear the latch holding bit
            _iEdgeCnt      := 0;                                       // 清探针沿计数 / Probe edge counter cleared
            _iOutsideCnt   := 0;                                       // 清窗口外计数 / Out-of-window counter cleared
            _eState        := E_DL_MeasureInputLatch_State.eIdle;       // 回空闲相，不滞留故障态 / Back to idle, never parked in fault
        END_IF

ELSE
    (* 迁移⑨（枚举兜底）：非法枚举值 → 故障级 99（R6） *)
    IF NOT _bFaultLatch THEN
        _iErrLatch   := 99;                    // 故障级：非法状态枚举值 / Fault: illegal state enum value
        _bFaultLatch := TRUE;                  // 置故障锁存（码位赋值 3 行内配对，R45）/ Latch the fault within three lines
    END_IF
END_CASE

(* —— 段 7：当拍故障请求锁存（域闸）+ 段尾迁移闸 + 撤使能降级（R191 已声明为降级+置标志） —— *)
IF (NOT _bCfgOk) AND (NOT _bFaultLatch) THEN
    _iErrLatch   := _iErrTmp;                  // 锁存域闸首因 / Latch the gate first cause
    _bFaultLatch := TRUE;                      // 置故障锁存 / Latch the fault
END_IF
IF _bFaultReq AND (NOT _bFaultLatch) THEN
    _iErrLatch   := _iErrTmp;                  // 锁存布防超时首因 / Latch the arming timeout cause
    _bFaultLatch := TRUE;                      // 置故障锁存 / Latch the fault
END_IF
IF _bFaultLatch AND (_eState <> E_DL_MeasureInputLatch_State.eFault) THEN
    _eState := E_DL_MeasureInputLatch_State.eFault;   // 锁存即迁相（段尾统一执行，FB50-1④）/ Latch forces the fault phase at the tail
END_IF
IF (NOT bEnable) AND (NOT _bFaultLatch) AND (_eState <> E_DL_MeasureInputLatch_State.eIdle) THEN
    _bLatchedLatch := FALSE;                   // 撤使能：锁存位撤销（保留上次锁存位置事实）/ Disable: latch cleared, the last position fact is kept
    _eState        := E_DL_MeasureInputLatch_State.eIdle;   // 撤使能：回空闲相 / Disable: back to idle
END_IF

(* —— 段 8：统一出口（单点映射；连续量出口做非有限防护，FB51-3 / R273） —— *)
eState  := _eState;                            // 相位映射 / Phase mapping
bArmed  := (_eState = E_DL_MeasureInputLatch_State.eArmed);   // 布防中（仅布防相为真）/ Armed, true only inside the armed phase
bLatched := _bLatchedLatch AND (NOT _bFaultLatch);            // 锁存有效（故障期强制撤销）/ Latch valid, forced off during fault
bDone   := _bDonePulse AND (NOT _bFaultLatch);                // 完成单拍（故障期强制撤销）/ Completion pulse forced off during fault
bError  := _bFaultLatch;                       // 故障标志取锁存位 / Fault flag taken from the latch
IF _bFaultLatch THEN
    iErrCode := _iErrLatch;                    // 故障期回放锁存码（FB33-1）/ Replay the latched code during fault
ELSE
    iErrCode := 0;                             // 非故障拍错误码归零 / Error code zeroed outside fault
END_IF
IF (_fLatchPos <> _fLatchPos) OR ((_fLatchPos - _fLatchPos) <> (_fLatchPos - _fLatchPos)) THEN
    rLatchPosMm := 0.0;                        // 保持槽污染兜底：归零（连续量安全侧）/ Contaminated holding value forced to zero
ELSE
    rLatchPosMm := LREAL_TO_REAL(_fLatchPos);  // 锁存位置出口（降位为 REAL）/ Latched position outlet demoted to REAL
END_IF
iOutsideCnt := _iOutsideCnt;                   // 窗口外计数映射 / Out-of-window counter mapping
iEdgeCnt    := _iEdgeCnt;                      // 探针沿计数映射 / Probe edge counter mapping
END_FUNCTION_BLOCK
